screen "P_Bar_1" 1024x768
   Bar "Default" at 10,10 size 40x120
   TextField "Label_Default" at 10,132 size 51x20; Text 'Default'
   Bar "BackColor" at 60,10 size 40x120
   TextField "Label_BackColor" at 60,132 size 67x20; Text 'BackColor'
   Bar "BarBackColor" at 110,10 size 40x120
   TextField "Label_BarBackColor" at 110,132 size 89x20; Text 'BarBackColor'
   Bar "BarEdgeStyle" at 160,10 size 40x120
   TextField "Label_BarEdgeStyle" at 160,132 size 90x20; Text 'BarEdgeStyle'
   Bar "BarEdgeStyle_2" at 210,10 size 40x120
   TextField "Label_BarEdgeStyle_2" at 210,132 size 106x20; Text 'BarEdgeStyle_2'
   Bar "BarOrientation" at 260,10 size 40x120
   TextField "Label_BarOrientation" at 260,132 size 99x20; Text 'BarOrientation'
   Bar "BarOrientation_2" at 310,10 size 40x120
   TextField "Label_BarOrientation_2" at 310,132 size 115x20; Text 'BarOrientation_2'
   Bar "BarOrientation_3" at 360,10 size 40x120
   TextField "Label_BarOrientation_3" at 360,132 size 115x20; Text 'BarOrientation_3'
   Bar "BorderBackColor" at 410,10 size 40x120
   TextField "Label_BorderBackColor" at 410,132 size 111x20; Text 'BorderBackColor'
   Bar "BorderColor" at 460,10 size 40x120
   TextField "Label_BorderColor" at 460,132 size 81x20; Text 'BorderColor'
   Bar "BorderWidth" at 510,10 size 40x120
   TextField "Label_BorderWidth" at 510,132 size 86x20; Text 'BorderWidth'
   Bar "CornerRadius" at 560,10 size 40x120
   TextField "Label_CornerRadius" at 560,132 size 91x20; Text 'CornerRadius'
   Bar "CountSubDivisions" at 610,10 size 40x120
   TextField "Label_CountSubDivisions" at 610,132 size 122x20; Text 'CountSubDivisions'
   Bar "EdgeStyle" at 660,10 size 40x120
   TextField "Label_EdgeStyle" at 660,132 size 68x20; Text 'EdgeStyle'
   Bar "EdgeStyle_2" at 710,10 size 40x120
   TextField "Label_EdgeStyle_2" at 710,132 size 84x20; Text 'EdgeStyle_2'
   Bar "EdgeStyle_3" at 760,10 size 40x120
   TextField "Label_EdgeStyle_3" at 760,132 size 84x20; Text 'EdgeStyle_3'
   Bar "EdgeStyle_4" at 810,10 size 40x120
   TextField "Label_EdgeStyle_4" at 810,132 size 84x20; Text 'EdgeStyle_4'
   Bar "Flashing" at 860,10 size 40x120
   TextField "Label_Flashing" at 860,132 size 55x20; Text 'Flashing'
   Bar "FlashingOnLimitViolation" at 910,10 size 40x120
   TextField "Label_FlashingOnLimitViolation" at 910,132 size 158x20; Text 'FlashingOnLimitViolation'
   Bar "ForeColor" at 960,10 size 40x120
   TextField "Label_ForeColor" at 960,132 size 65x20; Text 'ForeColor'
   Bar "IntegerDigits" at 10,156 size 40x120
   TextField "Label_IntegerDigits" at 10,278 size 89x20; Text 'IntegerDigits'
   Bar "LargeTickLabelingStep" at 60,156 size 40x120
   TextField "Label_LargeTickLabelingStep" at 60,278 size 148x20; Text 'LargeTickLabelingStep'
   Bar "MaximumValue" at 110,156 size 40x120; MaximumValue 200
   TextField "Label_MaximumValue" at 110,278 size 99x20; Text 'MaximumValue'
   Bar "MinimumValue" at 160,156 size 40x120; MinimumValue -100
   TextField "Label_MinimumValue" at 160,278 size 95x20; Text 'MinimumValue'
   Bar "Precision" at 210,156 size 40x120
   TextField "Label_Precision" at 210,278 size 62x20; Text 'Precision'
   Bar "RangeLower1Color" at 260,156 size 40x120
   TextField "Label_RangeLower1Color" at 260,278 size 126x20; Text 'RangeLower1Color'
   Bar "RangeLower1Enabled" at 310,156 size 40x120
   TextField "Label_RangeLower1Enabled" at 310,278 size 143x20; Text 'RangeLower1Enabled'
   Bar "RangeLower2Color" at 360,156 size 40x120
   TextField "Label_RangeLower2Color" at 360,278 size 126x20; Text 'RangeLower2Color'
   Bar "RangeLower2Enabled" at 410,156 size 40x120
   TextField "Label_RangeLower2Enabled" at 410,278 size 143x20; Text 'RangeLower2Enabled'
   Bar "RangeNormalColor" at 460,156 size 40x120
   TextField "Label_RangeNormalColor" at 460,278 size 122x20; Text 'RangeNormalColor'
   Bar "RangeNormalEnabled" at 510,156 size 40x120
   TextField "Label_RangeNormalEnabled" at 510,278 size 139x20; Text 'RangeNormalEnabled'
   Bar "RangeUpper1Color" at 560,156 size 40x120
   TextField "Label_RangeUpper1Color" at 560,278 size 124x20; Text 'RangeUpper1Color'
   Bar "RangeUpper1Enabled" at 610,156 size 40x120
   TextField "Label_RangeUpper1Enabled" at 610,278 size 141x20; Text 'RangeUpper1Enabled'
   Bar "RangeUpper2Color" at 660,156 size 40x120
   TextField "Label_RangeUpper2Color" at 660,278 size 124x20; Text 'RangeUpper2Color'
   Bar "RangeUpper2Enabled" at 710,156 size 40x120
   TextField "Label_RangeUpper2Enabled" at 710,278 size 141x20; Text 'RangeUpper2Enabled'
   Bar "ScaleColor" at 760,156 size 40x120
   TextField "Label_ScaleColor" at 760,278 size 71x20; Text 'ScaleColor'
   Bar "ScaleGradation" at 810,156 size 40x120
   TextField "Label_ScaleGradation" at 810,278 size 101x20; Text 'ScaleGradation'
   Bar "ScaleLabelingDoubleLined" at 860,156 size 40x120
   TextField "Label_ScaleLabelingDoubleLined" at 860,278 size 169x20; Text 'ScaleLabelingDoubleLined'
   Bar "ScalePosition" at 910,156 size 40x120
   TextField "Label_ScalePosition" at 910,278 size 89x20; Text 'ScalePosition'
   Bar "SegmentColoring" at 960,156 size 40x120
   TextField "Label_SegmentColoring" at 960,278 size 113x20; Text 'SegmentColoring'
   Bar "ShowLimitLines" at 10,302 size 40x120
   TextField "Label_ShowLimitLines" at 10,424 size 102x20; Text 'ShowLimitLines'
   Bar "ShowLimitMarkers" at 60,302 size 40x120
   TextField "Label_ShowLimitMarkers" at 60,424 size 122x20; Text 'ShowLimitMarkers'
   Bar "ShowLimitRanges" at 110,302 size 40x120
   TextField "Label_ShowLimitRanges" at 110,424 size 117x20; Text 'ShowLimitRanges'
   Bar "ShowProcessValue" at 160,302 size 40x120
   TextField "Label_ShowProcessValue" at 160,424 size 126x20; Text 'ShowProcessValue'
   Bar "ShowScale" at 210,302 size 40x120
   TextField "Label_ShowScale" at 210,424 size 73x20; Text 'ShowScale'
   Bar "ShowTickLabels" at 260,302 size 40x120
   TextField "Label_ShowTickLabels" at 260,424 size 104x20; Text 'ShowTickLabels'
   Bar "Unit" at 310,302 size 40x120; Unit mm
   TextField "Label_Unit" at 310,424 size 29x20; Text 'Unit'
   Bar "UseAutoScaling" at 360,302 size 40x120
   TextField "Label_UseAutoScaling" at 360,424 size 104x20; Text 'UseAutoScaling'
   Bar "UseDesignColorSchema" at 410,302 size 40x120
   TextField "Label_UseDesignColorSchema" at 410,424 size 153x20; Text 'UseDesignColorSchema'
   Bar "UseExponentialFormat" at 460,302 size 40x120
   TextField "Label_UseExponentialFormat" at 460,424 size 146x20; Text 'UseExponentialFormat'
   Button "Next" at 982,744 size 40x22; TextOff 'Text'
      on Click: ActivateScreen("P_Switch_1", 0)

screen "P_Switch_1" 1024x768
   Switch "Default" at 10,10 size 120x40; CaptionText 'Switch'; TextOff '0'; TextOn '1'
   TextField "Label_Default" at 10,52 size 51x20; Text 'Default'
   Switch "AboveUpperLimitColor" at 140,10 size 120x40; CaptionText 'Switch'; TextOff '0'; TextOn '1'
   TextField "Label_AboveUpperLimitColor" at 140,52 size 147x20; Text 'AboveUpperLimitColor'
   Switch "BackColor" at 270,10 size 120x40; CaptionText 'Switch'; TextOff '0'; TextOn '1'
   TextField "Label_BackColor" at 270,52 size 67x20; Text 'BackColor'
   Switch "BackFillStyle" at 400,10 size 120x40; CaptionText 'Switch'; TextOff '0'; TextOn '1'
   TextField "Label_BackFillStyle" at 400,52 size 82x20; Text 'BackFillStyle'
   Switch "BelowLowerLimitColor" at 530,10 size 120x40; CaptionText 'Switch'; TextOff '0'; TextOn '1'
   TextField "Label_BelowLowerLimitColor" at 530,52 size 145x20; Text 'BelowLowerLimitColor'
   Switch "BorderBackColor" at 660,10 size 120x40; CaptionText 'Switch'; TextOff '0'; TextOn '1'
   TextField "Label_BorderBackColor" at 660,52 size 111x20; Text 'BorderBackColor'
   Switch "BorderColor" at 790,10 size 120x40; CaptionText 'Switch'; TextOff '0'; TextOn '1'
   TextField "Label_BorderColor" at 790,52 size 81x20; Text 'BorderColor'
   Switch "BorderWidth" at 10,76 size 120x40; CaptionText 'Switch'; TextOff '0'; TextOn '1'
   TextField "Label_BorderWidth" at 10,118 size 86x20; Text 'BorderWidth'
   Switch "CaptionColor" at 140,76 size 120x40; CaptionText 'Switch'; TextOff '0'; TextOn '1'
   TextField "Label_CaptionColor" at 140,118 size 86x20; Text 'CaptionColor'
   Switch "CornerRadius" at 270,76 size 120x40; CaptionText 'Switch'; TextOff '0'; TextOn '1'
   TextField "Label_CornerRadius" at 270,118 size 91x20; Text 'CornerRadius'
   Switch "EdgeStyle" at 400,76 size 120x40; CaptionText 'Switch'; TextOff '0'; TextOn '1'
   TextField "Label_EdgeStyle" at 400,118 size 68x20; Text 'EdgeStyle'
   Switch "EdgeStyle_2" at 530,76 size 120x40; CaptionText 'Switch'; TextOff '0'; TextOn '1'
   TextField "Label_EdgeStyle_2" at 530,118 size 84x20; Text 'EdgeStyle_2'
   Switch "EdgeStyle_3" at 660,76 size 120x40; CaptionText 'Switch'; TextOff '0'; TextOn '1'
   TextField "Label_EdgeStyle_3" at 660,118 size 84x20; Text 'EdgeStyle_3'
   Switch "EdgeStyle_4" at 790,76 size 120x40; CaptionText 'Switch'; TextOff '0'; TextOn '1'
   TextField "Label_EdgeStyle_4" at 790,118 size 84x20; Text 'EdgeStyle_4'
   Switch "FirstGradientColor" at 10,142 size 120x40; CaptionText 'Switch'; TextOff '0'; TextOn '1'
   TextField "Label_FirstGradientColor" at 10,184 size 120x20; Text 'FirstGradientColor'
   Switch "FirstGradientOffset" at 140,142 size 120x40; CaptionText 'Switch'; TextOff '0'; TextOn '1'
   TextField "Label_FirstGradientOffset" at 140,184 size 127x20; Text 'FirstGradientOffset'
   Switch "FitToLargest" at 270,142 size 120x40; CaptionText 'Switch'; TextOff '0'; TextOn '1'
   TextField "Label_FitToLargest" at 270,184 size 84x20; Text 'FitToLargest'
   Switch "Flashing" at 400,142 size 120x40; CaptionText 'Switch'; TextOff '0'; TextOn '1'
   TextField "Label_Flashing" at 400,184 size 55x20; Text 'Flashing'
   Switch "FlashingOnLimitViolation" at 530,142 size 120x40; CaptionText 'Switch'; TextOff '0'; TextOn '1'
   TextField "Label_FlashingOnLimitViolation" at 530,184 size 158x20; Text 'FlashingOnLimitViolation'
   Switch "FocusColor" at 660,142 size 120x40; CaptionText 'Switch'; TextOff '0'; TextOn '1'
   TextField "Label_FocusColor" at 660,184 size 73x20; Text 'FocusColor'
   Switch "FocusWidth" at 790,142 size 120x40; CaptionText 'Switch'; TextOff '0'; TextOn '1'
   TextField "Label_FocusWidth" at 790,184 size 78x20; Text 'FocusWidth'
   Switch "ForeColor" at 10,208 size 120x40; CaptionText 'Switch'; TextOff '0'; TextOn '1'
   TextField "Label_ForeColor" at 10,250 size 65x20; Text 'ForeColor'
   Switch "HorizontalAlignment" at 140,208 size 120x40; CaptionText 'Switch'; TextOff '0'; TextOn '1'
   TextField "Label_HorizontalAlignment" at 140,250 size 135x20; Text 'HorizontalAlignment'
   Switch "HorizontalAlignment_2" at 270,208 size 120x40; CaptionText 'Switch'; TextOff '0'; TextOn '1'
   TextField "Label_HorizontalAlignment_2" at 270,250 size 151x20; Text 'HorizontalAlignment_2'
   Switch "HorizontalPictureAlignment" at 400,208 size 120x40; CaptionText 'Switch'; TextOff '0'; TextOn '1'
   TextField "Label_HorizontalPictureAlignment" at 400,250 size 181x20; Text 'HorizontalPictureAlignment'
   Switch "HorizontalPictureAlignment_2" at 530,208 size 120x40; CaptionText 'Switch'; TextOff '0'; TextOn '1'
   TextField "Label_HorizontalPictureAlignment_2" at 530,250 size 197x20; Text 'HorizontalPictureAlignment_2'
   Switch "InnerBackColorOff" at 660,208 size 120x40; CaptionText 'Switch'; TextOff '0'; TextOn '1'
   TextField "Label_InnerBackColorOff" at 660,250 size 121x20; Text 'InnerBackColorOff'
   Switch "InnerBackColorOn" at 790,208 size 120x40; CaptionText 'Switch'; TextOff '0'; TextOn '1'
   TextField "Label_InnerBackColorOn" at 790,250 size 119x20; Text 'InnerBackColorOn'
   Switch "MiddleGradientColor" at 10,274 size 120x40; CaptionText 'Switch'; TextOff '0'; TextOn '1'
   TextField "Label_MiddleGradientColor" at 10,316 size 133x20; Text 'MiddleGradientColor'
   Switch "PictureAreaBottomMargin" at 140,274 size 120x40; CaptionText 'Switch'; TextOff '0'; TextOn '1'
   TextField "Label_PictureAreaBottomMargin" at 140,316 size 173x20; Text 'PictureAreaBottomMargin'
   Switch "PictureAreaLeftMargin" at 270,274 size 120x40; CaptionText 'Switch'; TextOff '0'; TextOn '1'
   TextField "Label_PictureAreaLeftMargin" at 270,316 size 152x20; Text 'PictureAreaLeftMargin'
   Switch "PictureAreaRightMargin" at 400,274 size 120x40; CaptionText 'Switch'; TextOff '0'; TextOn '1'
   TextField "Label_PictureAreaRightMargin" at 400,316 size 160x20; Text 'PictureAreaRightMargin'
   Switch "PictureAreaTopMargin" at 530,274 size 120x40; CaptionText 'Switch'; TextOff '0'; TextOn '1'
   TextField "Label_PictureAreaTopMargin" at 530,316 size 149x20; Text 'PictureAreaTopMargin'
   Switch "SecondGradientColor" at 660,274 size 120x40; CaptionText 'Switch'; TextOff '0'; TextOn '1'
   TextField "Label_SecondGradientColor" at 660,316 size 139x20; Text 'SecondGradientColor'
   Switch "SecondGradientOffset" at 790,274 size 120x40; CaptionText 'Switch'; TextOff '0'; TextOn '1'
   TextField "Label_SecondGradientOffset" at 790,316 size 146x20; Text 'SecondGradientOffset'
   Switch "ShowCaption" at 10,340 size 120x40; CaptionText 'Switch'; TextOff '0'; TextOn '1'
   TextField "Label_ShowCaption" at 10,382 size 88x20; Text 'ShowCaption'
   Switch "SwitchOrientation" at 140,340 size 120x40; CaptionText 'Switch'; TextOff '0'; TextOn '1'
   TextField "Label_SwitchOrientation" at 140,382 size 120x20; Text 'SwitchOrientation'
   Switch "SwitchOrientation_2" at 270,340 size 120x40; CaptionText 'Switch'; TextOff '0'; TextOn '1'
   TextField "Label_SwitchOrientation_2" at 270,382 size 136x20; Text 'SwitchOrientation_2'
   Switch "SwitchOrientation_3" at 400,340 size 120x40; CaptionText 'Switch'; TextOff '0'; TextOn '1'
   TextField "Label_SwitchOrientation_3" at 400,382 size 136x20; Text 'SwitchOrientation_3'
   Switch "TextAreaBottomMargin" at 530,340 size 120x40; CaptionText 'Switch'; TextOff '0'; TextOn '1'
   TextField "Label_TextAreaBottomMargin" at 530,382 size 155x20; Text 'TextAreaBottomMargin'
   Switch "TextAreaLeftMargin" at 660,340 size 120x40; CaptionText 'Switch'; TextOff '0'; TextOn '1'
   TextField "Label_TextAreaLeftMargin" at 660,382 size 134x20; Text 'TextAreaLeftMargin'
   Switch "TextAreaRightMargin" at 790,340 size 120x40; CaptionText 'Switch'; TextOff '0'; TextOn '1'
   TextField "Label_TextAreaRightMargin" at 790,382 size 142x20; Text 'TextAreaRightMargin'
   Switch "TextAreaTopMargin" at 10,406 size 120x40; CaptionText 'Switch'; TextOff '0'; TextOn '1'
   TextField "Label_TextAreaTopMargin" at 10,448 size 131x20; Text 'TextAreaTopMargin'
   Switch "UseDesignColorSchema" at 140,406 size 120x40; CaptionText 'Switch'; TextOff '0'; TextOn '1'
   TextField "Label_UseDesignColorSchema" at 140,448 size 153x20; Text 'UseDesignColorSchema'
   Switch "UseFirstGradient" at 270,406 size 120x40; CaptionText 'Switch'; TextOff '0'; TextOn '1'
   TextField "Label_UseFirstGradient" at 270,448 size 110x20; Text 'UseFirstGradient'
   Switch "UseSecondGradient" at 400,406 size 120x40; CaptionText 'Switch'; TextOff '0'; TextOn '1'
   TextField "Label_UseSecondGradient" at 400,448 size 129x20; Text 'UseSecondGradient'
   Switch "VerticalAlignment" at 530,406 size 120x40; CaptionText 'Switch'; TextOff '0'; TextOn '1'
   TextField "Label_VerticalAlignment" at 530,448 size 119x20; Text 'VerticalAlignment'
   Switch "VerticalAlignment_2" at 660,406 size 120x40; CaptionText 'Switch'; TextOff '0'; TextOn '1'
   TextField "Label_VerticalAlignment_2" at 660,448 size 135x20; Text 'VerticalAlignment_2'
   Switch "VerticalPictureAlignment" at 790,406 size 120x40; CaptionText 'Switch'; TextOff '0'; TextOn '1'
   TextField "Label_VerticalPictureAlignment" at 790,448 size 165x20; Text 'VerticalPictureAlignment'
   Switch "VerticalPictureAlignment_2" at 10,472 size 120x40; CaptionText 'Switch'; TextOff '0'; TextOn '1'
   TextField "Label_VerticalPictureAlignment_2" at 10,514 size 181x20; Text 'VerticalPictureAlignment_2'
   Button "Next" at 982,744 size 40x22; TextOff 'Text'
      on Click: ActivateScreen("P_SymbolLibrary_1", 0)

screen "P_SymbolLibrary_1" 1024x768
   SymbolLibrary "Default" at 10,10 size 60x60
   TextField "Label_Default" at 10,72 size 51x20; Text 'Default'
   SymbolLibrary "AboveUpperLimitColor" at 80,10 size 60x60
   TextField "Label_AboveUpperLimitColor" at 80,72 size 147x20; Text 'AboveUpperLimitColor'
   SymbolLibrary "BackColor" at 150,10 size 60x60
   TextField "Label_BackColor" at 150,72 size 67x20; Text 'BackColor'
   SymbolLibrary "BackFillStyle" at 220,10 size 60x60
   TextField "Label_BackFillStyle" at 220,72 size 82x20; Text 'BackFillStyle'
   SymbolLibrary "BelowLowerLimitColor" at 290,10 size 60x60
   TextField "Label_BelowLowerLimitColor" at 290,72 size 145x20; Text 'BelowLowerLimitColor'
   SymbolLibrary "BlinkColor" at 360,10 size 60x60
   TextField "Label_BlinkColor" at 360,72 size 66x20; Text 'BlinkColor'
   SymbolLibrary "FillColorMode" at 430,10 size 60x60
   TextField "Label_FillColorMode" at 430,72 size 87x20; Text 'FillColorMode'
   SymbolLibrary "FillColorMode_2" at 500,10 size 60x60
   TextField "Label_FillColorMode_2" at 500,72 size 103x20; Text 'FillColorMode_2'
   SymbolLibrary "FixedAspectRatio" at 570,10 size 60x60
   TextField "Label_FixedAspectRatio" at 570,72 size 116x20; Text 'FixedAspectRatio'
   SymbolLibrary "Flashing" at 640,10 size 60x60
   TextField "Label_Flashing" at 640,72 size 55x20; Text 'Flashing'
   SymbolLibrary "FlashingOnLimitViolation" at 710,10 size 60x60
   TextField "Label_FlashingOnLimitViolation" at 710,72 size 158x20; Text 'FlashingOnLimitViolation'
   SymbolLibrary "Flip" at 780,10 size 60x60
   TextField "Label_Flip" at 780,72 size 24x20; Text 'Flip'
   SymbolLibrary "Flip_2" at 850,10 size 60x60
   TextField "Label_Flip_2" at 850,72 size 40x20; Text 'Flip_2'
   SymbolLibrary "Flip_3" at 920,10 size 60x60
   TextField "Label_Flip_3" at 920,72 size 40x20; Text 'Flip_3'
   SymbolLibrary "ForeColor" at 10,96 size 60x60
   TextField "Label_ForeColor" at 10,158 size 65x20; Text 'ForeColor'
   SymbolLibrary "Rotation" at 80,96 size 60x60
   TextField "Label_Rotation" at 80,158 size 60x20; Text 'Rotation'
   SymbolLibrary "Rotation_2" at 150,96 size 60x60
   TextField "Label_Rotation_2" at 150,158 size 76x20; Text 'Rotation_2'
   SymbolLibrary "Rotation_3" at 220,96 size 60x60
   TextField "Label_Rotation_3" at 220,158 size 76x20; Text 'Rotation_3'
   Button "Next" at 982,744 size 40x22; TextOff 'Text'
      on Click: ActivateScreen("P_Slider_1", 0)

screen "P_Slider_1" 1024x768
   Slider "Default" at 10,10 size 60x160; Caption 'SIMATIC'
   TextField "Label_Default" at 10,172 size 51x20; Text 'Default'
   Slider "BackColor" at 80,10 size 60x160; Caption 'SIMATIC'
   TextField "Label_BackColor" at 80,172 size 67x20; Text 'BackColor'
   Slider "BackFillStyle" at 150,10 size 60x160; Caption 'SIMATIC'
   TextField "Label_BackFillStyle" at 150,172 size 82x20; Text 'BackFillStyle'
   Slider "BarBackColor" at 220,10 size 60x160; Caption 'SIMATIC'
   TextField "Label_BarBackColor" at 220,172 size 89x20; Text 'BarBackColor'
   Slider "BarColor" at 290,10 size 60x160; Caption 'SIMATIC'
   TextField "Label_BarColor" at 290,172 size 59x20; Text 'BarColor'
   Slider "BarOrientation" at 360,10 size 60x160; Caption 'SIMATIC'
   TextField "Label_BarOrientation" at 360,172 size 99x20; Text 'BarOrientation'
   Slider "BarOrientation_2" at 430,10 size 60x160; Caption 'SIMATIC'
   TextField "Label_BarOrientation_2" at 430,172 size 115x20; Text 'BarOrientation_2'
   Slider "BarOrientation_3" at 500,10 size 60x160; Caption 'SIMATIC'
   TextField "Label_BarOrientation_3" at 500,172 size 115x20; Text 'BarOrientation_3'
   Slider "BorderBackColor" at 570,10 size 60x160; Caption 'SIMATIC'
   TextField "Label_BorderBackColor" at 570,172 size 111x20; Text 'BorderBackColor'
   Slider "BorderBrightColor3D" at 640,10 size 60x160; Caption 'SIMATIC'
   TextField "Label_BorderBrightColor3D" at 640,172 size 137x20; Text 'BorderBrightColor3D'
   Slider "BorderColor" at 710,10 size 60x160; Caption 'SIMATIC'
   TextField "Label_BorderColor" at 710,172 size 81x20; Text 'BorderColor'
   Slider "BorderInnerStyle3D" at 780,10 size 60x160; Caption 'SIMATIC'
   TextField "Label_BorderInnerStyle3D" at 780,172 size 133x20; Text 'BorderInnerStyle3D'
   Slider "BorderInnerStyle3D_2" at 850,10 size 60x160; Caption 'SIMATIC'
   TextField "Label_BorderInnerStyle3D_2" at 850,172 size 149x20; Text 'BorderInnerStyle3D_2'
   Slider "BorderInnerWidth3D" at 920,10 size 60x160; Caption 'SIMATIC'
   TextField "Label_BorderInnerWidth3D" at 920,172 size 138x20; Text 'BorderInnerWidth3D'
   Slider "BorderOuterStyle3D" at 10,196 size 60x160; Caption 'SIMATIC'
   TextField "Label_BorderOuterStyle3D" at 10,358 size 135x20; Text 'BorderOuterStyle3D'
   Slider "BorderOuterStyle3D_2" at 80,196 size 60x160; Caption 'SIMATIC'
   TextField "Label_BorderOuterStyle3D_2" at 80,358 size 151x20; Text 'BorderOuterStyle3D_2'
   Slider "BorderOuterWidth3D" at 150,196 size 60x160; Caption 'SIMATIC'
   TextField "Label_BorderOuterWidth3D" at 150,358 size 140x20; Text 'BorderOuterWidth3D'
   Slider "BorderShadeColor3D" at 220,196 size 60x160; Caption 'SIMATIC'
   TextField "Label_BorderShadeColor3D" at 220,358 size 138x20; Text 'BorderShadeColor3D'
   Slider "BorderWidth" at 290,196 size 60x160; Caption 'SIMATIC'
   TextField "Label_BorderWidth" at 290,358 size 86x20; Text 'BorderWidth'
   Slider "CornerRadius" at 360,196 size 60x160; Caption 'SIMATIC'
   TextField "Label_CornerRadius" at 360,358 size 91x20; Text 'CornerRadius'
   Slider "EdgeStyle" at 430,196 size 60x160; Caption 'SIMATIC'
   TextField "Label_EdgeStyle" at 430,358 size 68x20; Text 'EdgeStyle'
   Slider "EdgeStyle_2" at 500,196 size 60x160; Caption 'SIMATIC'
   TextField "Label_EdgeStyle_2" at 500,358 size 84x20; Text 'EdgeStyle_2'
   Slider "EdgeStyle_3" at 570,196 size 60x160; Caption 'SIMATIC'
   TextField "Label_EdgeStyle_3" at 570,358 size 84x20; Text 'EdgeStyle_3'
   Slider "EdgeStyle_4" at 640,196 size 60x160; Caption 'SIMATIC'
   TextField "Label_EdgeStyle_4" at 640,358 size 84x20; Text 'EdgeStyle_4'
   Slider "Flashing" at 710,196 size 60x160; Caption 'SIMATIC'
   TextField "Label_Flashing" at 710,358 size 55x20; Text 'Flashing'
   Slider "FocusColor" at 780,196 size 60x160; Caption 'SIMATIC'
   TextField "Label_FocusColor" at 780,358 size 73x20; Text 'FocusColor'
   Slider "FocusWidth" at 850,196 size 60x160; Caption 'SIMATIC'
   TextField "Label_FocusWidth" at 850,358 size 78x20; Text 'FocusWidth'
   Slider "ForeColor" at 920,196 size 60x160; Caption 'SIMATIC'
   TextField "Label_ForeColor" at 920,358 size 65x20; Text 'ForeColor'
   Slider "LabelColor" at 10,382 size 60x160; Caption 'SIMATIC'
   TextField "Label_LabelColor" at 10,544 size 71x20; Text 'LabelColor'
   Slider "MaximumValue" at 80,382 size 60x160; Caption 'SIMATIC'
   TextField "Label_MaximumValue" at 80,544 size 99x20; Text 'MaximumValue'
   Slider "MinimumValue" at 150,382 size 60x160; Caption 'SIMATIC'
   TextField "Label_MinimumValue" at 150,544 size 95x20; Text 'MinimumValue'
   Slider "RangeLower1Color" at 220,382 size 60x160; Caption 'SIMATIC'
   TextField "Label_RangeLower1Color" at 220,544 size 126x20; Text 'RangeLower1Color'
   Slider "RangeLower1Enabled" at 290,382 size 60x160; Caption 'SIMATIC'
   TextField "Label_RangeLower1Enabled" at 290,544 size 143x20; Text 'RangeLower1Enabled'
   Slider "RangeLower2Color" at 360,382 size 60x160; Caption 'SIMATIC'
   TextField "Label_RangeLower2Color" at 360,544 size 126x20; Text 'RangeLower2Color'
   Slider "RangeLower2Enabled" at 430,382 size 60x160; Caption 'SIMATIC'
   TextField "Label_RangeLower2Enabled" at 430,544 size 143x20; Text 'RangeLower2Enabled'
   Slider "RangeNormalColor" at 500,382 size 60x160; Caption 'SIMATIC'
   TextField "Label_RangeNormalColor" at 500,544 size 122x20; Text 'RangeNormalColor'
   Slider "RangeNormalEnabled" at 570,382 size 60x160; Caption 'SIMATIC'
   TextField "Label_RangeNormalEnabled" at 570,544 size 139x20; Text 'RangeNormalEnabled'
   Slider "RangeUpper1Color" at 640,382 size 60x160; Caption 'SIMATIC'
   TextField "Label_RangeUpper1Color" at 640,544 size 124x20; Text 'RangeUpper1Color'
   Slider "RangeUpper1Enabled" at 710,382 size 60x160; Caption 'SIMATIC'
   TextField "Label_RangeUpper1Enabled" at 710,544 size 141x20; Text 'RangeUpper1Enabled'
   Slider "RangeUpper2Color" at 780,382 size 60x160; Caption 'SIMATIC'
   TextField "Label_RangeUpper2Color" at 780,544 size 124x20; Text 'RangeUpper2Color'
   Slider "RangeUpper2Enabled" at 850,382 size 60x160; Caption 'SIMATIC'
   TextField "Label_RangeUpper2Enabled" at 850,544 size 141x20; Text 'RangeUpper2Enabled'
   Slider "ScalePosition" at 920,382 size 60x160; Caption 'SIMATIC'
   TextField "Label_ScalePosition" at 920,544 size 89x20; Text 'ScalePosition'
   Button "Next" at 982,744 size 40x22; TextOff 'Text'
      on Click: ActivateScreen("P_Slider_2", 0)

screen "P_Slider_2" 1024x768
   Slider "ShowBar" at 10,10 size 60x160; Caption 'SIMATIC'
   TextField "Label_ShowBar" at 10,172 size 61x20; Text 'ShowBar'
   Slider "ShowLimitLines" at 80,10 size 60x160; Caption 'SIMATIC'
   TextField "Label_ShowLimitLines" at 80,172 size 102x20; Text 'ShowLimitLines'
   Slider "ShowLimitMarkers" at 150,10 size 60x160; Caption 'SIMATIC'
   TextField "Label_ShowLimitMarkers" at 150,172 size 122x20; Text 'ShowLimitMarkers'
   Slider "ShowLimitRanges" at 220,10 size 60x160; Caption 'SIMATIC'
   TextField "Label_ShowLimitRanges" at 220,172 size 117x20; Text 'ShowLimitRanges'
   Slider "ShowPosition" at 290,10 size 60x160; Caption 'SIMATIC'
   TextField "Label_ShowPosition" at 290,172 size 90x20; Text 'ShowPosition'
   Slider "ShowScale" at 360,10 size 60x160; Caption 'SIMATIC'
   TextField "Label_ShowScale" at 360,172 size 73x20; Text 'ShowScale'
   Slider "ShowThumb" at 430,10 size 60x160; Caption 'SIMATIC'
   TextField "Label_ShowThumb" at 430,172 size 81x20; Text 'ShowThumb'
   Slider "ShowTickLabels" at 500,10 size 60x160; Caption 'SIMATIC'
   TextField "Label_ShowTickLabels" at 500,172 size 104x20; Text 'ShowTickLabels'
   Slider "ShowTicks" at 570,10 size 60x160; Caption 'SIMATIC'
   TextField "Label_ShowTicks" at 570,172 size 70x20; Text 'ShowTicks'
   Slider "ThumbBackColor" at 640,10 size 60x160; Caption 'SIMATIC'
   TextField "Label_ThumbBackColor" at 640,172 size 109x20; Text 'ThumbBackColor'
   Slider "UseDesignColorSchema" at 710,10 size 60x160; Caption 'SIMATIC'
   TextField "Label_UseDesignColorSchema" at 710,172 size 153x20; Text 'UseDesignColorSchema'
   Button "Next" at 982,744 size 40x22; TextOff 'Text'
      on Click: ActivateScreen("P_Gauge_1", 0)

screen "P_Gauge_1" 1024x768
   Gauge "Default" at 10,10 size 150x150; CaptionText 'SIMATIC'
   TextField "Label_Default" at 10,162 size 51x20; Text 'Default'
   Gauge "AngleMax" at 170,10 size 150x150; CaptionText 'SIMATIC'
   TextField "Label_AngleMax" at 170,162 size 67x20; Text 'AngleMax'
   Gauge "AngleMin" at 330,10 size 150x150; CaptionText 'SIMATIC'
   TextField "Label_AngleMin" at 330,162 size 63x20; Text 'AngleMin'
   Gauge "BackColor" at 490,10 size 150x150; CaptionText 'SIMATIC'
   TextField "Label_BackColor" at 490,162 size 67x20; Text 'BackColor'
   Gauge "BackFillStyle" at 650,10 size 150x150; CaptionText 'SIMATIC'
   TextField "Label_BackFillStyle" at 650,162 size 82x20; Text 'BackFillStyle'
   Gauge "BorderBackColor" at 810,10 size 150x150; CaptionText 'SIMATIC'
   TextField "Label_BorderBackColor" at 810,162 size 111x20; Text 'BorderBackColor'
   Gauge "BorderColor" at 10,186 size 150x150; CaptionText 'SIMATIC'
   TextField "Label_BorderColor" at 10,338 size 81x20; Text 'BorderColor'
   Gauge "BorderWidth" at 170,186 size 150x150; CaptionText 'SIMATIC'
   TextField "Label_BorderWidth" at 170,338 size 86x20; Text 'BorderWidth'
   Gauge "CaptionColor" at 330,186 size 150x150; CaptionText 'SIMATIC'
   TextField "Label_CaptionColor" at 330,338 size 86x20; Text 'CaptionColor'
   Gauge "CaptionTop" at 490,186 size 150x150; CaptionText 'SIMATIC'
   TextField "Label_CaptionTop" at 490,338 size 76x20; Text 'CaptionTop'
   Gauge "CenterColor" at 650,186 size 150x150; CaptionText 'SIMATIC'
   TextField "Label_CenterColor" at 650,338 size 81x20; Text 'CenterColor'
   Gauge "CenterSize" at 810,186 size 150x150; CaptionText 'SIMATIC'
   TextField "Label_CenterSize" at 810,338 size 74x20; Text 'CenterSize'
   Gauge "CornerRadius" at 10,362 size 150x150; CaptionText 'SIMATIC'
   TextField "Label_CornerRadius" at 10,514 size 91x20; Text 'CornerRadius'
   Gauge "DialColor" at 170,362 size 150x150; CaptionText 'SIMATIC'
   TextField "Label_DialColor" at 170,514 size 60x20; Text 'DialColor'
   Gauge "DialFillStyle" at 330,362 size 150x150; CaptionText 'SIMATIC'
   TextField "Label_DialFillStyle" at 330,514 size 75x20; Text 'DialFillStyle'
   Gauge "DialSize" at 490,362 size 150x150; CaptionText 'SIMATIC'
   TextField "Label_DialSize" at 490,514 size 53x20; Text 'DialSize'
   Gauge "EdgeStyle" at 650,362 size 150x150; CaptionText 'SIMATIC'
   TextField "Label_EdgeStyle" at 650,514 size 68x20; Text 'EdgeStyle'
   Gauge "EdgeStyle_2" at 810,362 size 150x150; CaptionText 'SIMATIC'
   TextField "Label_EdgeStyle_2" at 810,514 size 84x20; Text 'EdgeStyle_2'
   Gauge "EdgeStyle_3" at 10,538 size 150x150; CaptionText 'SIMATIC'
   TextField "Label_EdgeStyle_3" at 10,690 size 84x20; Text 'EdgeStyle_3'
   Gauge "EdgeStyle_4" at 170,538 size 150x150; CaptionText 'SIMATIC'
   TextField "Label_EdgeStyle_4" at 170,690 size 84x20; Text 'EdgeStyle_4'
   Gauge "Gradation" at 330,538 size 150x150; CaptionText 'SIMATIC'
   TextField "Label_Gradation" at 330,690 size 67x20; Text 'Gradation'
   Gauge "InnerDialColor" at 490,538 size 150x150; CaptionText 'SIMATIC'
   TextField "Label_InnerDialColor" at 490,690 size 95x20; Text 'InnerDialColor'
   Gauge "InnerDialInnerDistance" at 650,538 size 150x150; CaptionText 'SIMATIC'
   TextField "Label_InnerDialInnerDistance" at 650,690 size 153x20; Text 'InnerDialInnerDistance'
   Gauge "InnerDialOuterDistance" at 810,538 size 150x150; CaptionText 'SIMATIC'
   TextField "Label_InnerDialOuterDistance" at 810,690 size 155x20; Text 'InnerDialOuterDistance'
   Button "Next" at 982,744 size 40x22; TextOff 'Text'
      on Click: ActivateScreen("P_Gauge_2", 0)

screen "P_Gauge_2" 1024x768
   Gauge "LockSquaredExtent" at 10,10 size 150x150; CaptionText 'SIMATIC'
   TextField "Label_LockSquaredExtent" at 10,162 size 129x20; Text 'LockSquaredExtent'
   Gauge "MaximumValue" at 170,10 size 150x150; CaptionText 'SIMATIC'
   TextField "Label_MaximumValue" at 170,162 size 99x20; Text 'MaximumValue'
   Gauge "MinimumValue" at 330,10 size 150x150; CaptionText 'SIMATIC'
   TextField "Label_MinimumValue" at 330,162 size 95x20; Text 'MinimumValue'
   Gauge "NeedleHeight" at 490,10 size 150x150; CaptionText 'SIMATIC'
   TextField "Label_NeedleHeight" at 490,162 size 89x20; Text 'NeedleHeight'
   Gauge "PointerColor" at 650,10 size 150x150; CaptionText 'SIMATIC'
   TextField "Label_PointerColor" at 650,162 size 84x20; Text 'PointerColor'
   Gauge "RangeLower1Color" at 810,10 size 150x150; CaptionText 'SIMATIC'
   TextField "Label_RangeLower1Color" at 810,162 size 126x20; Text 'RangeLower1Color'
   Gauge "RangeLower1Enabled" at 10,186 size 150x150; CaptionText 'SIMATIC'
   TextField "Label_RangeLower1Enabled" at 10,338 size 143x20; Text 'RangeLower1Enabled'
   Gauge "RangeLower2Color" at 170,186 size 150x150; CaptionText 'SIMATIC'
   TextField "Label_RangeLower2Color" at 170,338 size 126x20; Text 'RangeLower2Color'
   Gauge "RangeLower2Enabled" at 330,186 size 150x150; CaptionText 'SIMATIC'
   TextField "Label_RangeLower2Enabled" at 330,338 size 143x20; Text 'RangeLower2Enabled'
   Gauge "RangeNormalColor" at 490,186 size 150x150; CaptionText 'SIMATIC'
   TextField "Label_RangeNormalColor" at 490,338 size 122x20; Text 'RangeNormalColor'
   Gauge "RangeNormalEnabled" at 650,186 size 150x150; CaptionText 'SIMATIC'
   TextField "Label_RangeNormalEnabled" at 650,338 size 139x20; Text 'RangeNormalEnabled'
   Gauge "RangeUpper1Color" at 810,186 size 150x150; CaptionText 'SIMATIC'
   TextField "Label_RangeUpper1Color" at 810,338 size 124x20; Text 'RangeUpper1Color'
   Gauge "RangeUpper1Enabled" at 10,362 size 150x150; CaptionText 'SIMATIC'
   TextField "Label_RangeUpper1Enabled" at 10,514 size 141x20; Text 'RangeUpper1Enabled'
   Gauge "RangeUpper1Start" at 170,362 size 150x150; CaptionText 'SIMATIC'
   TextField "Label_RangeUpper1Start" at 170,514 size 125x20; Text 'RangeUpper1Start'
   Gauge "RangeUpper2Color" at 330,362 size 150x150; CaptionText 'SIMATIC'
   TextField "Label_RangeUpper2Color" at 330,514 size 124x20; Text 'RangeUpper2Color'
   Gauge "RangeUpper2Enabled" at 490,362 size 150x150; CaptionText 'SIMATIC'
   TextField "Label_RangeUpper2Enabled" at 490,514 size 141x20; Text 'RangeUpper2Enabled'
   Gauge "RangeUpper2Start" at 650,362 size 150x150; CaptionText 'SIMATIC'
   TextField "Label_RangeUpper2Start" at 650,514 size 125x20; Text 'RangeUpper2Start'
   Gauge "ScaleLabelColor" at 810,362 size 150x150; CaptionText 'SIMATIC'
   TextField "Label_ScaleLabelColor" at 810,514 size 105x20; Text 'ScaleLabelColor'
   Gauge "ScaleTickColor" at 10,538 size 150x150; CaptionText 'SIMATIC'
   TextField "Label_ScaleTickColor" at 10,690 size 95x20; Text 'ScaleTickColor'
   Gauge "ScaleTickLabelPosition" at 170,538 size 150x150; CaptionText 'SIMATIC'
   TextField "Label_ScaleTickLabelPosition" at 170,690 size 147x20; Text 'ScaleTickLabelPosition'
   Gauge "ScaleTickLength" at 330,538 size 150x150; CaptionText 'SIMATIC'
   TextField "Label_ScaleTickLength" at 330,690 size 107x20; Text 'ScaleTickLength'
   Gauge "ScaleTickPosition" at 490,538 size 150x150; CaptionText 'SIMATIC'
   TextField "Label_ScaleTickPosition" at 490,690 size 113x20; Text 'ScaleTickPosition'
   Gauge "ShowDecimalPoint" at 650,538 size 150x150; CaptionText 'SIMATIC'
   TextField "Label_ShowDecimalPoint" at 650,690 size 121x20; Text 'ShowDecimalPoint'
   Gauge "ShowInnerDial" at 810,538 size 150x150; CaptionText 'SIMATIC'
   TextField "Label_ShowInnerDial" at 810,690 size 97x20; Text 'ShowInnerDial'
   Button "Next" at 982,744 size 40x22; TextOff 'Text'
      on Click: ActivateScreen("P_Gauge_3", 0)

screen "P_Gauge_3" 1024x768
   Gauge "ShowLimitRanges" at 10,10 size 150x150; CaptionText 'SIMATIC'
   TextField "Label_ShowLimitRanges" at 10,162 size 117x20; Text 'ShowLimitRanges'
   Gauge "ShowPeakValuePointer" at 170,10 size 150x150; CaptionText 'SIMATIC'
   TextField "Label_ShowPeakValuePointer" at 170,162 size 153x20; Text 'ShowPeakValuePointer'
   Gauge "UnitColor" at 330,10 size 150x150; CaptionText 'SIMATIC'
   TextField "Label_UnitColor" at 330,162 size 62x20; Text 'UnitColor'
   Gauge "UnitTop" at 490,10 size 150x150; CaptionText 'SIMATIC'
   TextField "Label_UnitTop" at 490,162 size 52x20; Text 'UnitTop'
   Gauge "UseDesignColorSchema" at 650,10 size 150x150; CaptionText 'SIMATIC'
   TextField "Label_UseDesignColorSchema" at 650,162 size 153x20; Text 'UseDesignColorSchema'
   Button "Next" at 982,744 size 40x22; TextOff 'Text'
      on Click: ActivateScreen("P_Clock_1", 0)

screen "P_Clock_1" 1024x768
   Clock "Default" at 10,10 size 150x150
   TextField "Label_Default" at 10,162 size 51x20; Text 'Default'
   Clock "Analog" at 170,10 size 150x150
   TextField "Label_Analog" at 170,162 size 49x20; Text 'Analog'
   Clock "BackFillStyle" at 330,10 size 150x150
   TextField "Label_BackFillStyle" at 330,162 size 82x20; Text 'BackFillStyle'
   Clock "BorderBackColor" at 490,10 size 150x150
   TextField "Label_BorderBackColor" at 490,162 size 111x20; Text 'BorderBackColor'
   Clock "BorderColor" at 650,10 size 150x150
   TextField "Label_BorderColor" at 650,162 size 81x20; Text 'BorderColor'
   Clock "BorderWidth" at 810,10 size 150x150
   TextField "Label_BorderWidth" at 810,162 size 86x20; Text 'BorderWidth'
   Clock "CornerRadius" at 10,186 size 150x150
   TextField "Label_CornerRadius" at 10,338 size 91x20; Text 'CornerRadius'
   Clock "DialColor" at 170,186 size 150x150
   TextField "Label_DialColor" at 170,338 size 60x20; Text 'DialColor'
   Clock "EdgeStyle" at 330,186 size 150x150
   TextField "Label_EdgeStyle" at 330,338 size 68x20; Text 'EdgeStyle'
   Clock "EdgeStyle_2" at 490,186 size 150x150
   TextField "Label_EdgeStyle_2" at 490,338 size 84x20; Text 'EdgeStyle_2'
   Clock "EdgeStyle_3" at 650,186 size 150x150
   TextField "Label_EdgeStyle_3" at 650,338 size 84x20; Text 'EdgeStyle_3'
   Clock "EdgeStyle_4" at 810,186 size 150x150
   TextField "Label_EdgeStyle_4" at 810,338 size 84x20; Text 'EdgeStyle_4'
   Clock "Flashing" at 10,362 size 150x150
   TextField "Label_Flashing" at 10,514 size 55x20; Text 'Flashing'
   Clock "HourNeedleHeight" at 170,362 size 150x150
   TextField "Label_HourNeedleHeight" at 170,514 size 120x20; Text 'HourNeedleHeight'
   Clock "HourNeedleWidth" at 330,362 size 150x150
   TextField "Label_HourNeedleWidth" at 330,514 size 116x20; Text 'HourNeedleWidth'
   Clock "LockSquaredExtent" at 490,362 size 150x150
   TextField "Label_LockSquaredExtent" at 490,514 size 129x20; Text 'LockSquaredExtent'
   Clock "MinuteNeedleHeight" at 650,362 size 150x150
   TextField "Label_MinuteNeedleHeight" at 650,514 size 133x20; Text 'MinuteNeedleHeight'
   Clock "MinuteNeedleWidth" at 810,362 size 150x150
   TextField "Label_MinuteNeedleWidth" at 810,514 size 129x20; Text 'MinuteNeedleWidth'
   Clock "NeedleBorderColor" at 10,538 size 150x150
   TextField "Label_NeedleBorderColor" at 10,690 size 124x20; Text 'NeedleBorderColor'
   Clock "NeedleColor" at 170,538 size 150x150
   TextField "Label_NeedleColor" at 170,690 size 80x20; Text 'NeedleColor'
   Clock "NeedleFillStyle" at 330,538 size 150x150
   TextField "Label_NeedleFillStyle" at 330,690 size 95x20; Text 'NeedleFillStyle'
   Clock "NumberStyle" at 490,538 size 150x150
   TextField "Label_NumberStyle" at 490,690 size 86x20; Text 'NumberStyle'
   Clock "NumberStyle_2" at 650,538 size 150x150
   TextField "Label_NumberStyle_2" at 650,690 size 102x20; Text 'NumberStyle_2'
   Clock "SecondNeedleHeight" at 810,538 size 150x150
   TextField "Label_SecondNeedleHeight" at 810,690 size 136x20; Text 'SecondNeedleHeight'
   Button "Next" at 982,744 size 40x22; TextOff 'Text'
      on Click: ActivateScreen("P_Clock_2", 0)

screen "P_Clock_2" 1024x768
   Clock "SecondNeedleWidth" at 10,10 size 150x150
   TextField "Label_SecondNeedleWidth" at 10,162 size 132x20; Text 'SecondNeedleWidth'
   Clock "ShowTicks" at 170,10 size 150x150
   TextField "Label_ShowTicks" at 170,162 size 70x20; Text 'ShowTicks'
   Clock "TickDistance" at 330,10 size 150x150
   TextField "Label_TickDistance" at 330,162 size 84x20; Text 'TickDistance'
   Clock "TickStyle" at 490,10 size 150x150
   TextField "Label_TickStyle" at 490,162 size 61x20; Text 'TickStyle'
   Clock "TicksColor" at 650,10 size 150x150
   TextField "Label_TicksColor" at 650,162 size 68x20; Text 'TicksColor'
   Clock "UseDesignColorSchema" at 810,10 size 150x150
   TextField "Label_UseDesignColorSchema" at 810,162 size 153x20; Text 'UseDesignColorSchema'
   Button "Next" at 982,744 size 40x22; TextOff 'Text'
      on Click: ActivateScreen("P_Line_1", 0)

screen "P_IOField_1" 1024x768
   IOField "Default" at 10,10 size 100x30
   TextField "Label_Default" at 10,42 size 51x20; Text 'Default'
   IOField "AboveUpperLimitColor" at 120,10 size 100x30
   TextField "Label_AboveUpperLimitColor" at 120,42 size 147x20; Text 'AboveUpperLimitColor'
   IOField "BackColor" at 230,10 size 100x30
   TextField "Label_BackColor" at 230,42 size 67x20; Text 'BackColor'
   IOField "BackFillStyle" at 340,10 size 100x30
   TextField "Label_BackFillStyle" at 340,42 size 82x20; Text 'BackFillStyle'
   IOField "BelowLowerLimitColor" at 450,10 size 100x30
   TextField "Label_BelowLowerLimitColor" at 450,42 size 145x20; Text 'BelowLowerLimitColor'
   IOField "BorderBackColor" at 560,10 size 100x30
   TextField "Label_BorderBackColor" at 560,42 size 111x20; Text 'BorderBackColor'
   IOField "BorderColor" at 670,10 size 100x30
   TextField "Label_BorderColor" at 670,42 size 81x20; Text 'BorderColor'
   IOField "BorderWidth" at 780,10 size 100x30
   TextField "Label_BorderWidth" at 780,42 size 86x20; Text 'BorderWidth'
   IOField "BottomMargin" at 890,10 size 100x30
   TextField "Label_BottomMargin" at 890,42 size 95x20; Text 'BottomMargin'
   IOField "CornerRadius" at 10,66 size 100x30
   TextField "Label_CornerRadius" at 10,98 size 91x20; Text 'CornerRadius'
   IOField "DataFormat_3" at 120,66 size 100x30
   TextField "Label_DataFormat_3" at 120,98 size 96x20; Text 'DataFormat_3'
   IOField "EdgeStyle" at 230,66 size 100x30
   TextField "Label_EdgeStyle" at 230,98 size 68x20; Text 'EdgeStyle'
   IOField "EdgeStyle_2" at 340,66 size 100x30
   TextField "Label_EdgeStyle_2" at 340,98 size 84x20; Text 'EdgeStyle_2'
   IOField "EdgeStyle_3" at 450,66 size 100x30
   TextField "Label_EdgeStyle_3" at 450,98 size 84x20; Text 'EdgeStyle_3'
   IOField "EdgeStyle_4" at 560,66 size 100x30
   TextField "Label_EdgeStyle_4" at 560,98 size 84x20; Text 'EdgeStyle_4'
   IOField "FieldLength" at 670,66 size 100x30
   TextField "Label_FieldLength" at 670,98 size 77x20; Text 'FieldLength'
   IOField "FitToLargest" at 780,66 size 75x30
   TextField "Label_FitToLargest" at 780,98 size 84x20; Text 'FitToLargest'
   IOField "Flashing" at 890,66 size 100x30
   TextField "Label_Flashing" at 890,98 size 55x20; Text 'Flashing'
   IOField "ForeColor" at 10,122 size 100x30
   TextField "Label_ForeColor" at 10,154 size 65x20; Text 'ForeColor'
   IOField "FormatPattern" at 120,122 size 100x30; FormatPattern 99.9
   TextField "Label_FormatPattern" at 120,154 size 99x20; Text 'FormatPattern'
   IOField "HorizontalAlignment" at 230,122 size 100x30
   TextField "Label_HorizontalAlignment" at 230,154 size 135x20; Text 'HorizontalAlignment'
   IOField "HorizontalAlignment_2" at 340,122 size 100x30
   TextField "Label_HorizontalAlignment_2" at 340,154 size 151x20; Text 'HorizontalAlignment_2'
   IOField "LeftMargin" at 450,122 size 100x30
   TextField "Label_LeftMargin" at 450,154 size 74x20; Text 'LeftMargin'
   IOField "Mode" at 560,122 size 100x30
   TextField "Label_Mode" at 560,154 size 39x20; Text 'Mode'
   IOField "Mode_2" at 670,122 size 100x30
   TextField "Label_Mode_2" at 670,154 size 55x20; Text 'Mode_2'
   IOField "RightMargin" at 780,122 size 100x30
   TextField "Label_RightMargin" at 780,154 size 82x20; Text 'RightMargin'
   IOField "ShiftDecimalPoint" at 890,122 size 100x30
   TextField "Label_ShiftDecimalPoint" at 890,154 size 116x20; Text 'ShiftDecimalPoint'
   IOField "ShowLeadingZeros" at 10,178 size 100x30
   TextField "Label_ShowLeadingZeros" at 10,210 size 125x20; Text 'ShowLeadingZeros'
   IOField "TopMargin" at 120,178 size 100x30
   TextField "Label_TopMargin" at 120,210 size 71x20; Text 'TopMargin'
   IOField "Unit" at 230,178 size 100x30; Unit mm
   TextField "Label_Unit" at 230,210 size 29x20; Text 'Unit'
   IOField "UseDesignColorSchema" at 340,178 size 100x30
   TextField "Label_UseDesignColorSchema" at 340,210 size 153x20; Text 'UseDesignColorSchema'
   IOField "VerticalAlignment" at 450,178 size 100x30
   TextField "Label_VerticalAlignment" at 450,210 size 119x20; Text 'VerticalAlignment'
   IOField "VerticalAlignment_2" at 560,178 size 100x30
   TextField "Label_VerticalAlignment_2" at 560,210 size 135x20; Text 'VerticalAlignment_2'
   Button "Next" at 982,744 size 40x22; TextOff 'Text'
      on Click: ActivateScreen("P_Button_1", 0)

screen "D_Bar_1" 1024x768
   Bar "Static" at 6,4 size 40x120
   TextField "Label_Static" at 6,156 size 42x20; Text 'Static'
   Bar "A_Range" at 98,4 size 40x120
      Appearance <- "D_Range"
   TextField "Label_A_Range" at 98,156 size 63x20; Text 'A_Range'
   Bar "A_Flash" at 190,4 size 40x120
      Appearance <- "D_Range"
   TextField "Label_A_Flash" at 190,156 size 54x20; Text 'A_Flash'
   Bar "A_Bit" at 282,4 size 40x120
      Appearance <- "D_Bool"
   TextField "Label_A_Bit" at 282,156 size 39x20; Text 'A_Bit'
   Bar "A_Bits" at 374,4 size 40x120
      Appearance <- "D_Bits"
   TextField "Label_A_Bits" at 374,156 size 46x20; Text 'A_Bits'
   Bar "V_Range" at 466,4 size 40x120
      Visibility <- "D_Range"
   TextField "Label_V_Range" at 466,156 size 62x20; Text 'V_Range'
   Bar "V_Bit" at 558,4 size 40x120
      Visibility <- "D_Vis"
   TextField "Label_V_Bit" at 558,156 size 38x20; Text 'V_Bit'
   Bar "M_H" at 650,4 size 40x120
      HorizontalMovement <- "D_Pct"
   TextField "Label_M_H" at 650,156 size 32x20; Text 'M_H'
   Bar "M_V" at 742,4 size 40x120
      VerticalMovement <- "D_Pct"
   TextField "Label_M_V" at 742,156 size 32x20; Text 'M_V'
   Bar "M_D" at 834,4 size 40x120
      DiagonalMovement <- "D_Pct"
   TextField "Label_M_D" at 834,156 size 32x20; Text 'M_D'
   Bar "M_Direct" at 926,4 size 40x120
      DirectMovement <- "D_X"
      DirectMovement <- "D_Y"
   TextField "Label_M_Direct" at 926,156 size 62x20; Text 'M_Direct'
   Bar "E_Range" at 6,176 size 40x120
      ObjectEnable <- "D_Range"
   TextField "Label_E_Range" at 6,328 size 60x20; Text 'E_Range'
   Bar "E_Bit" at 98,176 size 40x120
      ObjectEnable <- "D_En"
   TextField "Label_E_Bit" at 98,328 size 36x20; Text 'E_Bit'
   Bar "PV_Pct" at 190,176 size 40x120
      ProcessValue <- "D_Pct"
   TextField "Label_PV_Pct" at 190,328 size 50x20; Text 'PV_Pct'
   Bar "PV_Real" at 282,176 size 40x120
      ProcessValue <- "D_Real"
   TextField "Label_PV_Real" at 282,328 size 57x20; Text 'PV_Real'
   Bar "PV_BarR" at 374,176 size 40x120
      ProcessValue <- "D_BarR"
   TextField "Label_PV_BarR" at 374,328 size 60x20; Text 'PV_BarR'
   Bar "PV_Pct_0_100" at 466,176 size 40x120; MinimumValue 0; MaximumValue 100
      ProcessValue <- "D_Pct"
   TextField "Label_PV_Pct_0_100" at 466,328 size 98x20; Text 'PV_Pct_0_100'
   Bar "PV_Pct_MaxMin" at 558,176 size 40x120
      ProcessValue <- "D_Pct"
      MaximumValue <- "D_Max"
      MinimumValue <- "D_Min"
   TextField "Label_PV_Pct_MaxMin" at 558,328 size 106x20; Text 'PV_Pct_MaxMin'
   IOField "State" at 4,742 size 60x22; FormatPattern 9
      ProcessValue <- "D_State"
   Button "S1" at 70,742 size 40x22; TextOff 'S1'
      on Click: "SetS1"()
   Button "S2" at 114,742 size 40x22; TextOff 'S2'
      on Click: "SetS2"()
   Button "S3" at 158,742 size 40x22; TextOff 'S3'
      on Click: "SetS3"()
   Button "S4" at 202,742 size 40x22; TextOff 'S4'
      on Click: "SetS4"()
   Button "Next" at 980,742 size 40x22; TextOff 'Next'
      on Click: ActivateScreen("D_Switch_1", 0)

screen "D_Button_1" 1024x768
   Button "Static" at 6,4 size 100x40; TextOff 'Text'
   TextField "Label_Static" at 6,76 size 42x20; Text 'Static'
   Button "A_Range" at 158,4 size 100x40; TextOff 'Text'
      Appearance <- "D_Range"
   TextField "Label_A_Range" at 158,76 size 63x20; Text 'A_Range'
   Button "A_Flash" at 310,4 size 100x40; TextOff 'Text'
      Appearance <- "D_Range"
   TextField "Label_A_Flash" at 310,76 size 54x20; Text 'A_Flash'
   Button "A_Bit" at 462,4 size 100x40; TextOff 'Text'
      Appearance <- "D_Bool"
   TextField "Label_A_Bit" at 462,76 size 39x20; Text 'A_Bit'
   Button "A_Bits" at 614,4 size 100x40; TextOff 'Text'
      Appearance <- "D_Bits"
   TextField "Label_A_Bits" at 614,76 size 46x20; Text 'A_Bits'
   Button "V_Range" at 766,4 size 100x40; TextOff 'Text'
      Visibility <- "D_Range"
   TextField "Label_V_Range" at 766,76 size 62x20; Text 'V_Range'
   Button "V_Bit" at 6,96 size 100x40; TextOff 'Text'
      Visibility <- "D_Vis"
   TextField "Label_V_Bit" at 6,168 size 38x20; Text 'V_Bit'
   Button "M_H" at 158,96 size 100x40; TextOff 'Text'
      HorizontalMovement <- "D_Pct"
   TextField "Label_M_H" at 158,168 size 32x20; Text 'M_H'
   Button "M_V" at 310,96 size 100x40; TextOff 'Text'
      VerticalMovement <- "D_Pct"
   TextField "Label_M_V" at 310,168 size 32x20; Text 'M_V'
   Button "M_D" at 462,96 size 100x40; TextOff 'Text'
      DiagonalMovement <- "D_Pct"
   TextField "Label_M_D" at 462,168 size 32x20; Text 'M_D'
   Button "M_Direct" at 614,96 size 100x40; TextOff 'Text'
      DirectMovement <- "D_X"
      DirectMovement <- "D_Y"
   TextField "Label_M_Direct" at 614,168 size 62x20; Text 'M_Direct'
   Button "E_Range" at 766,96 size 100x40; TextOff 'Text'
      ObjectEnable <- "D_Range"
   TextField "Label_E_Range" at 766,168 size 60x20; Text 'E_Range'
   Button "E_Bit" at 6,188 size 100x40; TextOff 'Text'
      ObjectEnable <- "D_En"
   TextField "Label_E_Bit" at 6,260 size 36x20; Text 'E_Bit'
   IOField "State" at 4,742 size 60x22; FormatPattern 9
      ProcessValue <- "D_State"
   Button "S1" at 70,742 size 40x22; TextOff 'S1'
      on Click: "SetS1"()
   Button "S2" at 114,742 size 40x22; TextOff 'S2'
      on Click: "SetS2"()
   Button "S3" at 158,742 size 40x22; TextOff 'S3'
      on Click: "SetS3"()
   Button "S4" at 202,742 size 40x22; TextOff 'S4'
      on Click: "SetS4"()
   Button "Next" at 980,742 size 40x22; TextOff 'Next'
      on Click: ActivateScreen("D_SymbolicIOField_1", 0)

screen "D_Circle_1" 1024x768
   TextField "Label_Static" at 6,86 size 42x20; Text 'Static'
   Circle "A_Range" at 108,4 size 50x50
      Appearance <- "D_Range"
   TextField "Label_A_Range" at 108,86 size 63x20; Text 'A_Range'
   Circle "A_Flash" at 210,4 size 50x50
      Appearance <- "D_Range"
   TextField "Label_A_Flash" at 210,86 size 54x20; Text 'A_Flash'
   Circle "A_Bit" at 312,4 size 50x50
      Appearance <- "D_Bool"
   TextField "Label_A_Bit" at 312,86 size 39x20; Text 'A_Bit'
   Circle "A_Bits" at 414,4 size 50x50
      Appearance <- "D_Bits"
   TextField "Label_A_Bits" at 414,86 size 46x20; Text 'A_Bits'
   Circle "V_Range" at 516,4 size 50x50
      Visibility <- "D_Range"
   TextField "Label_V_Range" at 516,86 size 62x20; Text 'V_Range'
   Circle "V_Bit" at 618,4 size 50x50
      Visibility <- "D_Vis"
   TextField "Label_V_Bit" at 618,86 size 38x20; Text 'V_Bit'
   Circle "M_H" at 720,4 size 50x50
      HorizontalMovement <- "D_Pct"
   TextField "Label_M_H" at 720,86 size 32x20; Text 'M_H'
   Circle "M_V" at 822,4 size 50x50
      VerticalMovement <- "D_Pct"
   TextField "Label_M_V" at 822,86 size 32x20; Text 'M_V'
   Circle "M_D" at 6,106 size 50x50
      DiagonalMovement <- "D_Pct"
   TextField "Label_M_D" at 6,188 size 32x20; Text 'M_D'
   Circle "M_Direct" at 108,106 size 50x50
      DirectMovement <- "D_X"
      DirectMovement <- "D_Y"
   TextField "Label_M_Direct" at 108,188 size 62x20; Text 'M_Direct'
   Circle "E_Range" at 210,106 size 50x50
      ObjectEnable <- "D_Range"
   TextField "Label_E_Range" at 210,188 size 60x20; Text 'E_Range'
   Circle "E_Bit" at 312,106 size 50x50
      ObjectEnable <- "D_En"
   TextField "Label_E_Bit" at 312,188 size 36x20; Text 'E_Bit'
   IOField "State" at 4,742 size 60x22; FormatPattern 9
      ProcessValue <- "D_State"
   Button "S1" at 70,742 size 40x22; TextOff 'S1'
      on Click: "SetS1"()
   Button "S2" at 114,742 size 40x22; TextOff 'S2'
      on Click: "SetS2"()
   Button "S3" at 158,742 size 40x22; TextOff 'S3'
      on Click: "SetS3"()
   Button "S4" at 202,742 size 40x22; TextOff 'S4'
      on Click: "SetS4"()
   Button "Next" at 980,742 size 40x22; TextOff 'Next'
      on Click: ActivateScreen("D_Rectangle_1", 0)

screen "D_Clock_1" 1024x768
   Clock "Static" at 6,4 size 150x150
   TextField "Label_Static" at 6,186 size 42x20; Text 'Static'
   Clock "A_Range" at 208,4 size 150x150
      Appearance <- "D_Range"
   TextField "Label_A_Range" at 208,186 size 63x20; Text 'A_Range'
   Clock "A_Flash" at 410,4 size 150x150
      Appearance <- "D_Range"
   TextField "Label_A_Flash" at 410,186 size 54x20; Text 'A_Flash'
   Clock "A_Bit" at 612,4 size 150x150
      Appearance <- "D_Bool"
   TextField "Label_A_Bit" at 612,186 size 39x20; Text 'A_Bit'
   Clock "A_Bits" at 814,4 size 150x150
      Appearance <- "D_Bits"
   TextField "Label_A_Bits" at 814,186 size 46x20; Text 'A_Bits'
   Clock "V_Range" at 6,206 size 150x150
      Visibility <- "D_Range"
   TextField "Label_V_Range" at 6,388 size 62x20; Text 'V_Range'
   Clock "V_Bit" at 208,206 size 150x150
      Visibility <- "D_Vis"
   TextField "Label_V_Bit" at 208,388 size 38x20; Text 'V_Bit'
   Clock "M_H" at 410,206 size 150x150
      HorizontalMovement <- "D_Pct"
   TextField "Label_M_H" at 410,388 size 32x20; Text 'M_H'
   Clock "M_V" at 612,206 size 150x150
      VerticalMovement <- "D_Pct"
   TextField "Label_M_V" at 612,388 size 32x20; Text 'M_V'
   Clock "M_D" at 814,206 size 150x150
      DiagonalMovement <- "D_Pct"
   TextField "Label_M_D" at 814,388 size 32x20; Text 'M_D'
   Clock "M_Direct" at 6,408 size 150x150
      DirectMovement <- "D_X"
      DirectMovement <- "D_Y"
   TextField "Label_M_Direct" at 6,590 size 62x20; Text 'M_Direct'
   Clock "E_Range" at 208,408 size 150x150
      ObjectEnable <- "D_Range"
   TextField "Label_E_Range" at 208,590 size 60x20; Text 'E_Range'
   Clock "E_Bit" at 410,408 size 150x150
      ObjectEnable <- "D_En"
   TextField "Label_E_Bit" at 410,590 size 36x20; Text 'E_Bit'
   IOField "State" at 4,742 size 60x22; FormatPattern 9
      ProcessValue <- "D_State"
   Button "S1" at 70,742 size 40x22; TextOff 'S1'
      on Click: "SetS1"()
   Button "S2" at 114,742 size 40x22; TextOff 'S2'
      on Click: "SetS2"()
   Button "S3" at 158,742 size 40x22; TextOff 'S3'
      on Click: "SetS3"()
   Button "S4" at 202,742 size 40x22; TextOff 'S4'
      on Click: "SetS4"()
   Button "Next" at 980,742 size 40x22; TextOff 'Next'
      on Click: ActivateScreen("D_Line_1", 0)

screen "D_DateTimeField_1" 1024x768
   DateTimeField "Static" at 6,4 size 189x26
   TextField "Label_Static" at 6,66 size 42x20; Text 'Static'
   DateTimeField "A_Range" at 218,4 size 189x26
      Appearance <- "D_Range"
   TextField "Label_A_Range" at 218,66 size 63x20; Text 'A_Range'
   DateTimeField "A_Flash" at 430,4 size 189x26
      Appearance <- "D_Range"
   TextField "Label_A_Flash" at 430,66 size 54x20; Text 'A_Flash'
   DateTimeField "A_Bit" at 642,4 size 189x26
      Appearance <- "D_Bool"
   TextField "Label_A_Bit" at 642,66 size 39x20; Text 'A_Bit'
   DateTimeField "A_Bits" at 6,86 size 189x26
      Appearance <- "D_Bits"
   TextField "Label_A_Bits" at 6,148 size 46x20; Text 'A_Bits'
   DateTimeField "V_Range" at 218,86 size 189x26
      Visibility <- "D_Range"
   TextField "Label_V_Range" at 218,148 size 62x20; Text 'V_Range'
   DateTimeField "V_Bit" at 430,86 size 189x26
      Visibility <- "D_Vis"
   TextField "Label_V_Bit" at 430,148 size 38x20; Text 'V_Bit'
   DateTimeField "M_H" at 642,86 size 189x26
      HorizontalMovement <- "D_Pct"
   TextField "Label_M_H" at 642,148 size 32x20; Text 'M_H'
   DateTimeField "M_V" at 6,168 size 189x26
      VerticalMovement <- "D_Pct"
   TextField "Label_M_V" at 6,230 size 32x20; Text 'M_V'
   DateTimeField "M_D" at 218,168 size 189x26
      DiagonalMovement <- "D_Pct"
   TextField "Label_M_D" at 218,230 size 32x20; Text 'M_D'
   DateTimeField "M_Direct" at 430,168 size 189x26
      DirectMovement <- "D_X"
      DirectMovement <- "D_Y"
   TextField "Label_M_Direct" at 430,230 size 62x20; Text 'M_Direct'
   DateTimeField "E_Range" at 642,168 size 189x26
      ObjectEnable <- "D_Range"
   TextField "Label_E_Range" at 642,230 size 60x20; Text 'E_Range'
   DateTimeField "E_Bit" at 6,250 size 189x26
      ObjectEnable <- "D_En"
   TextField "Label_E_Bit" at 6,312 size 36x20; Text 'E_Bit'
   DateTimeField "PV_DateTime" at 218,250 size 189x26
      ProcessValue <- "D_DateTime"
   TextField "Label_PV_DateTime" at 218,312 size 89x20; Text 'PV_DateTime'
   IOField "State" at 4,742 size 60x22; FormatPattern 9
      ProcessValue <- "D_State"
   Button "S1" at 70,742 size 40x22; TextOff 'S1'
      on Click: "SetS1"()
   Button "S2" at 114,742 size 40x22; TextOff 'S2'
      on Click: "SetS2"()
   Button "S3" at 158,742 size 40x22; TextOff 'S3'
      on Click: "SetS3"()
   Button "S4" at 202,742 size 40x22; TextOff 'S4'
      on Click: "SetS4"()
   Button "Next" at 980,742 size 40x22; TextOff 'Next'
      on Click: ActivateScreen("D_Bar_1", 0)

screen "D_Ellipse_1" 1024x768
   TextField "Label_Static" at 6,86 size 42x20; Text 'Static'
   Ellipse "A_Range" at 158,4 size 100x50
      Appearance <- "D_Range"
   TextField "Label_A_Range" at 158,86 size 63x20; Text 'A_Range'
   Ellipse "A_Flash" at 310,4 size 100x50
      Appearance <- "D_Range"
   TextField "Label_A_Flash" at 310,86 size 54x20; Text 'A_Flash'
   Ellipse "A_Bit" at 462,4 size 100x50
      Appearance <- "D_Bool"
   TextField "Label_A_Bit" at 462,86 size 39x20; Text 'A_Bit'
   Ellipse "A_Bits" at 614,4 size 100x50
      Appearance <- "D_Bits"
   TextField "Label_A_Bits" at 614,86 size 46x20; Text 'A_Bits'
   Ellipse "V_Range" at 766,4 size 100x50
      Visibility <- "D_Range"
   TextField "Label_V_Range" at 766,86 size 62x20; Text 'V_Range'
   Ellipse "V_Bit" at 6,106 size 100x50
      Visibility <- "D_Vis"
   TextField "Label_V_Bit" at 6,188 size 38x20; Text 'V_Bit'
   Ellipse "M_H" at 158,106 size 100x50
      HorizontalMovement <- "D_Pct"
   TextField "Label_M_H" at 158,188 size 32x20; Text 'M_H'
   Ellipse "M_V" at 310,106 size 100x50
      VerticalMovement <- "D_Pct"
   TextField "Label_M_V" at 310,188 size 32x20; Text 'M_V'
   Ellipse "M_D" at 462,106 size 100x50
      DiagonalMovement <- "D_Pct"
   TextField "Label_M_D" at 462,188 size 32x20; Text 'M_D'
   Ellipse "M_Direct" at 614,106 size 100x50
      DirectMovement <- "D_X"
      DirectMovement <- "D_Y"
   TextField "Label_M_Direct" at 614,188 size 62x20; Text 'M_Direct'
   Ellipse "E_Range" at 766,106 size 100x50
      ObjectEnable <- "D_Range"
   TextField "Label_E_Range" at 766,188 size 60x20; Text 'E_Range'
   Ellipse "E_Bit" at 6,208 size 100x50
      ObjectEnable <- "D_En"
   TextField "Label_E_Bit" at 6,290 size 36x20; Text 'E_Bit'
   IOField "State" at 4,742 size 60x22; FormatPattern 9
      ProcessValue <- "D_State"
   Button "S1" at 70,742 size 40x22; TextOff 'S1'
      on Click: "SetS1"()
   Button "S2" at 114,742 size 40x22; TextOff 'S2'
      on Click: "SetS2"()
   Button "S3" at 158,742 size 40x22; TextOff 'S3'
      on Click: "SetS3"()
   Button "S4" at 202,742 size 40x22; TextOff 'S4'
      on Click: "SetS4"()
   Button "Next" at 980,742 size 40x22; TextOff 'Next'
      on Click: ActivateScreen("D_Circle_1", 0)

screen "D_Gauge_1" 1024x768
   Gauge "Static" at 6,4 size 150x150; CaptionText 'SIMATIC'
   TextField "Label_Static" at 6,186 size 42x20; Text 'Static'
   Gauge "A_Range" at 208,4 size 150x150; CaptionText 'SIMATIC'
      Appearance <- "D_Range"
   TextField "Label_A_Range" at 208,186 size 63x20; Text 'A_Range'
   Gauge "A_Flash" at 410,4 size 150x150; CaptionText 'SIMATIC'
      Appearance <- "D_Range"
   TextField "Label_A_Flash" at 410,186 size 54x20; Text 'A_Flash'
   Gauge "A_Bit" at 612,4 size 150x150; CaptionText 'SIMATIC'
      Appearance <- "D_Bool"
   TextField "Label_A_Bit" at 612,186 size 39x20; Text 'A_Bit'
   Gauge "A_Bits" at 814,4 size 150x150; CaptionText 'SIMATIC'
      Appearance <- "D_Bits"
   TextField "Label_A_Bits" at 814,186 size 46x20; Text 'A_Bits'
   Gauge "V_Range" at 6,206 size 150x150; CaptionText 'SIMATIC'
      Visibility <- "D_Range"
   TextField "Label_V_Range" at 6,388 size 62x20; Text 'V_Range'
   Gauge "V_Bit" at 208,206 size 150x150; CaptionText 'SIMATIC'
      Visibility <- "D_Vis"
   TextField "Label_V_Bit" at 208,388 size 38x20; Text 'V_Bit'
   Gauge "M_H" at 410,206 size 150x150; CaptionText 'SIMATIC'
      HorizontalMovement <- "D_Pct"
   TextField "Label_M_H" at 410,388 size 32x20; Text 'M_H'
   Gauge "M_V" at 612,206 size 150x150; CaptionText 'SIMATIC'
      VerticalMovement <- "D_Pct"
   TextField "Label_M_V" at 612,388 size 32x20; Text 'M_V'
   Gauge "M_D" at 814,206 size 150x150; CaptionText 'SIMATIC'
      DiagonalMovement <- "D_Pct"
   TextField "Label_M_D" at 814,388 size 32x20; Text 'M_D'
   Gauge "M_Direct" at 6,408 size 150x150; CaptionText 'SIMATIC'
      DirectMovement <- "D_X"
      DirectMovement <- "D_Y"
   TextField "Label_M_Direct" at 6,590 size 62x20; Text 'M_Direct'
   Gauge "E_Range" at 208,408 size 150x150; CaptionText 'SIMATIC'
      ObjectEnable <- "D_Range"
   TextField "Label_E_Range" at 208,590 size 60x20; Text 'E_Range'
   Gauge "E_Bit" at 410,408 size 150x150; CaptionText 'SIMATIC'
      ObjectEnable <- "D_En"
   TextField "Label_E_Bit" at 410,590 size 36x20; Text 'E_Bit'
   Gauge "PV_Pct" at 612,408 size 150x150; CaptionText 'SIMATIC'
      ProcessValue <- "D_Pct"
   TextField "Label_PV_Pct" at 612,590 size 50x20; Text 'PV_Pct'
   Gauge "PV_Real" at 814,408 size 150x150; CaptionText 'SIMATIC'
      ProcessValue <- "D_Real"
   TextField "Label_PV_Real" at 814,590 size 57x20; Text 'PV_Real'
   IOField "State" at 4,742 size 60x22; FormatPattern 9
      ProcessValue <- "D_State"
   Button "S1" at 70,742 size 40x22; TextOff 'S1'
      on Click: "SetS1"()
   Button "S2" at 114,742 size 40x22; TextOff 'S2'
      on Click: "SetS2"()
   Button "S3" at 158,742 size 40x22; TextOff 'S3'
      on Click: "SetS3"()
   Button "S4" at 202,742 size 40x22; TextOff 'S4'
      on Click: "SetS4"()
   Button "Next" at 980,742 size 40x22; TextOff 'Next'
      on Click: ActivateScreen("D_Gauge_2", 0)

screen "D_Gauge_2" 1024x768
   Gauge "PV_Pct_MaxMin" at 6,4 size 150x150; CaptionText 'SIMATIC'
      ProcessValue <- "D_Pct"
      MaximumValue <- "D_Max"
      MinimumValue <- "D_Min"
   TextField "Label_PV_Pct_MaxMin" at 6,186 size 106x20; Text 'PV_Pct_MaxMin'
   IOField "State" at 4,742 size 60x22; FormatPattern 9
      ProcessValue <- "D_State"
   Button "S1" at 70,742 size 40x22; TextOff 'S1'
      on Click: "SetS1"()
   Button "S2" at 114,742 size 40x22; TextOff 'S2'
      on Click: "SetS2"()
   Button "S3" at 158,742 size 40x22; TextOff 'S3'
      on Click: "SetS3"()
   Button "S4" at 202,742 size 40x22; TextOff 'S4'
      on Click: "SetS4"()
   Button "Next" at 980,742 size 40x22; TextOff 'Next'
      on Click: ActivateScreen("D_Clock_1", 0)

screen "D_GraphicIOField_1" 1024x768
   GraphicIOField "Static" at 6,4 size 60x60
   TextField "Label_Static" at 6,96 size 42x20; Text 'Static'
   GraphicIOField "A_Range" at 118,4 size 60x60
      Appearance <- "D_Range"
   TextField "Label_A_Range" at 118,96 size 63x20; Text 'A_Range'
   GraphicIOField "A_Flash" at 230,4 size 60x60
      Appearance <- "D_Range"
   TextField "Label_A_Flash" at 230,96 size 54x20; Text 'A_Flash'
   GraphicIOField "A_Bit" at 342,4 size 60x60
      Appearance <- "D_Bool"
   TextField "Label_A_Bit" at 342,96 size 39x20; Text 'A_Bit'
   GraphicIOField "A_Bits" at 454,4 size 60x60
      Appearance <- "D_Bits"
   TextField "Label_A_Bits" at 454,96 size 46x20; Text 'A_Bits'
   GraphicIOField "V_Range" at 566,4 size 60x60
      Visibility <- "D_Range"
   TextField "Label_V_Range" at 566,96 size 62x20; Text 'V_Range'
   GraphicIOField "V_Bit" at 678,4 size 60x60
      Visibility <- "D_Vis"
   TextField "Label_V_Bit" at 678,96 size 38x20; Text 'V_Bit'
   GraphicIOField "M_H" at 790,4 size 60x60
      HorizontalMovement <- "D_Pct"
   TextField "Label_M_H" at 790,96 size 32x20; Text 'M_H'
   GraphicIOField "M_V" at 902,4 size 60x60
      VerticalMovement <- "D_Pct"
   TextField "Label_M_V" at 902,96 size 32x20; Text 'M_V'
   GraphicIOField "M_D" at 6,116 size 60x60
      DiagonalMovement <- "D_Pct"
   TextField "Label_M_D" at 6,208 size 32x20; Text 'M_D'
   GraphicIOField "M_Direct" at 118,116 size 60x60
      DirectMovement <- "D_X"
      DirectMovement <- "D_Y"
   TextField "Label_M_Direct" at 118,208 size 62x20; Text 'M_Direct'
   GraphicIOField "E_Range" at 230,116 size 60x60
      ObjectEnable <- "D_Range"
   TextField "Label_E_Range" at 230,208 size 60x20; Text 'E_Range'
   GraphicIOField "E_Bit" at 342,116 size 60x60
      ObjectEnable <- "D_En"
   TextField "Label_E_Bit" at 342,208 size 36x20; Text 'E_Bit'
   IOField "State" at 4,742 size 60x22; FormatPattern 9
      ProcessValue <- "D_State"
   Button "S1" at 70,742 size 40x22; TextOff 'S1'
      on Click: "SetS1"()
   Button "S2" at 114,742 size 40x22; TextOff 'S2'
      on Click: "SetS2"()
   Button "S3" at 158,742 size 40x22; TextOff 'S3'
      on Click: "SetS3"()
   Button "S4" at 202,742 size 40x22; TextOff 'S4'
      on Click: "SetS4"()
   Button "Next" at 980,742 size 40x22; TextOff 'Next'
      on Click: ActivateScreen("D_DateTimeField_1", 0)

screen "D_GraphicView_1" 1024x768
   GraphicView "Static" at 6,4 size 100x60
   TextField "Label_Static" at 6,96 size 42x20; Text 'Static'
   GraphicView "A_Range" at 158,4 size 100x60
      Appearance <- "D_Range"
   TextField "Label_A_Range" at 158,96 size 63x20; Text 'A_Range'
   GraphicView "A_Flash" at 310,4 size 100x60
      Appearance <- "D_Range"
   TextField "Label_A_Flash" at 310,96 size 54x20; Text 'A_Flash'
   GraphicView "A_Bit" at 462,4 size 100x60
      Appearance <- "D_Bool"
   TextField "Label_A_Bit" at 462,96 size 39x20; Text 'A_Bit'
   GraphicView "A_Bits" at 614,4 size 100x60
      Appearance <- "D_Bits"
   TextField "Label_A_Bits" at 614,96 size 46x20; Text 'A_Bits'
   GraphicView "V_Range" at 766,4 size 100x60
      Visibility <- "D_Range"
   TextField "Label_V_Range" at 766,96 size 62x20; Text 'V_Range'
   GraphicView "V_Bit" at 6,116 size 100x60
      Visibility <- "D_Vis"
   TextField "Label_V_Bit" at 6,208 size 38x20; Text 'V_Bit'
   GraphicView "M_H" at 158,116 size 100x60
      HorizontalMovement <- "D_Pct"
   TextField "Label_M_H" at 158,208 size 32x20; Text 'M_H'
   GraphicView "M_V" at 310,116 size 100x60
      VerticalMovement <- "D_Pct"
   TextField "Label_M_V" at 310,208 size 32x20; Text 'M_V'
   GraphicView "M_D" at 462,116 size 100x60
      DiagonalMovement <- "D_Pct"
   TextField "Label_M_D" at 462,208 size 32x20; Text 'M_D'
   GraphicView "M_Direct" at 614,116 size 100x60
      DirectMovement <- "D_X"
      DirectMovement <- "D_Y"
   TextField "Label_M_Direct" at 614,208 size 62x20; Text 'M_Direct'
   GraphicView "E_Range" at 766,116 size 100x60
      ObjectEnable <- "D_Range"
   TextField "Label_E_Range" at 766,208 size 60x20; Text 'E_Range'
   GraphicView "E_Bit" at 6,228 size 100x60
      ObjectEnable <- "D_En"
   TextField "Label_E_Bit" at 6,320 size 36x20; Text 'E_Bit'
   IOField "State" at 4,742 size 60x22; FormatPattern 9
      ProcessValue <- "D_State"
   Button "S1" at 70,742 size 40x22; TextOff 'S1'
      on Click: "SetS1"()
   Button "S2" at 114,742 size 40x22; TextOff 'S2'
      on Click: "SetS2"()
   Button "S3" at 158,742 size 40x22; TextOff 'S3'
      on Click: "SetS3"()
   Button "S4" at 202,742 size 40x22; TextOff 'S4'
      on Click: "SetS4"()
   Button "Next" at 980,742 size 40x22; TextOff 'Next'
      on Click: ActivateScreen("D_IOField_1", 0)

screen "D_IOField_1" 1024x768
   IOField "Static" at 6,4 size 100x30
   TextField "Label_Static" at 6,66 size 42x20; Text 'Static'
   IOField "A_Range" at 158,4 size 100x30
      Appearance <- "D_Range"
   TextField "Label_A_Range" at 158,66 size 63x20; Text 'A_Range'
   IOField "A_Flash" at 310,4 size 100x30
      Appearance <- "D_Range"
   TextField "Label_A_Flash" at 310,66 size 54x20; Text 'A_Flash'
   IOField "A_Bit" at 462,4 size 100x30
      Appearance <- "D_Bool"
   TextField "Label_A_Bit" at 462,66 size 39x20; Text 'A_Bit'
   IOField "A_Bits" at 614,4 size 100x30
      Appearance <- "D_Bits"
   TextField "Label_A_Bits" at 614,66 size 46x20; Text 'A_Bits'
   IOField "V_Range" at 766,4 size 100x30
      Visibility <- "D_Range"
   TextField "Label_V_Range" at 766,66 size 62x20; Text 'V_Range'
   IOField "V_Bit" at 6,86 size 100x30
      Visibility <- "D_Vis"
   TextField "Label_V_Bit" at 6,148 size 38x20; Text 'V_Bit'
   IOField "M_H" at 158,86 size 100x30
      HorizontalMovement <- "D_Pct"
   TextField "Label_M_H" at 158,148 size 32x20; Text 'M_H'
   IOField "M_V" at 310,86 size 100x30
      VerticalMovement <- "D_Pct"
   TextField "Label_M_V" at 310,148 size 32x20; Text 'M_V'
   IOField "M_D" at 462,86 size 100x30
      DiagonalMovement <- "D_Pct"
   TextField "Label_M_D" at 462,148 size 32x20; Text 'M_D'
   IOField "M_Direct" at 614,86 size 100x30
      DirectMovement <- "D_X"
      DirectMovement <- "D_Y"
   TextField "Label_M_Direct" at 614,148 size 62x20; Text 'M_Direct'
   IOField "E_Range" at 766,86 size 100x30
      ObjectEnable <- "D_Range"
   TextField "Label_E_Range" at 766,148 size 60x20; Text 'E_Range'
   IOField "E_Bit" at 6,168 size 100x30
      ObjectEnable <- "D_En"
   TextField "Label_E_Bit" at 6,230 size 36x20; Text 'E_Bit'
   IOField "PV_SInt" at 158,168 size 100x30; FormatPattern s999
      ProcessValue <- "D_SInt"
   TextField "Label_PV_SInt" at 158,230 size 56x20; Text 'PV_SInt'
   IOField "PV_Int" at 310,168 size 100x30; FormatPattern s99999
      ProcessValue <- "D_Int"
   TextField "Label_PV_Int" at 310,230 size 48x20; Text 'PV_Int'
   IOField "PV_DInt" at 462,168 size 100x30; FormatPattern s9999999999
      ProcessValue <- "D_DInt"
   TextField "Label_PV_DInt" at 462,230 size 57x20; Text 'PV_DInt'
   IOField "PV_USInt" at 614,168 size 100x30; FormatPattern 999
      ProcessValue <- "D_USInt"
   TextField "Label_PV_USInt" at 614,230 size 64x20; Text 'PV_USInt'
   IOField "PV_UInt" at 766,168 size 100x30; FormatPattern 99999
      ProcessValue <- "D_UInt"
   TextField "Label_PV_UInt" at 766,230 size 56x20; Text 'PV_UInt'
   IOField "PV_UDInt" at 6,250 size 100x30; FormatPattern 9999999999
      ProcessValue <- "D_UDInt"
   TextField "Label_PV_UDInt" at 6,312 size 65x20; Text 'PV_UDInt'
   IOField "PV_Real" at 158,250 size 100x30
      ProcessValue <- "D_Real"
   TextField "Label_PV_Real" at 158,312 size 57x20; Text 'PV_Real'
   IOField "PV_LReal" at 310,250 size 100x30
      ProcessValue <- "D_LReal"
   TextField "Label_PV_LReal" at 310,312 size 64x20; Text 'PV_LReal'
   IOField "PV_String" at 462,250 size 100x30
      ProcessValue <- "D_String"
   TextField "Label_PV_String" at 462,312 size 68x20; Text 'PV_String'
   IOField "PV_Int_Shift2" at 614,250 size 100x30; FormatPattern s99999
      ProcessValue <- "D_Int"
   TextField "Label_PV_Int_Shift2" at 614,312 size 94x20; Text 'PV_Int_Shift2'
   IOField "PV_Int_s999999" at 766,250 size 100x30; FormatPattern s999999
      ProcessValue <- "D_Int"
   TextField "Label_PV_Int_s999999" at 766,312 size 111x20; Text 'PV_Int_s999999'
   IOField "PV_Real_s9999_99" at 6,332 size 100x30; FormatPattern s9999.99
      ProcessValue <- "D_Real"
   TextField "Label_PV_Real_s9999_99" at 6,394 size 128x20; Text 'PV_Real_s9999_99'
   IOField "PV_Int_Output" at 158,332 size 100x30; FormatPattern s99999
      ProcessValue <- "D_Int"
   TextField "Label_PV_Int_Output" at 158,394 size 101x20; Text 'PV_Int_Output'
   IOField "PV_Int_s99" at 310,332 size 100x30; FormatPattern s99
      ProcessValue <- "D_Int"
   TextField "Label_PV_Int_s99" at 310,394 size 79x20; Text 'PV_Int_s99'
   IOField "State" at 4,742 size 60x22; FormatPattern 9
      ProcessValue <- "D_State"
   Button "S1" at 70,742 size 40x22; TextOff 'S1'
      on Click: "SetS1"()
   Button "S2" at 114,742 size 40x22; TextOff 'S2'
      on Click: "SetS2"()
   Button "S3" at 158,742 size 40x22; TextOff 'S3'
      on Click: "SetS3"()
   Button "S4" at 202,742 size 40x22; TextOff 'S4'
      on Click: "SetS4"()
   Button "Next" at 980,742 size 40x22; TextOff 'Next'
      on Click: ActivateScreen("D_Button_1", 0)

screen "D_Line_1" 1024x768
   TextField "Label_Static" at 6,86 size 42x20; Text 'Static'
   Line "A_Range" at 158,4 size 100x50
      Appearance <- "D_Range"
   TextField "Label_A_Range" at 158,86 size 63x20; Text 'A_Range'
   Line "A_Flash" at 310,4 size 100x50
      Appearance <- "D_Range"
   TextField "Label_A_Flash" at 310,86 size 54x20; Text 'A_Flash'
   Line "A_Bit" at 462,4 size 100x50
      Appearance <- "D_Bool"
   TextField "Label_A_Bit" at 462,86 size 39x20; Text 'A_Bit'
   Line "A_Bits" at 614,4 size 100x50
      Appearance <- "D_Bits"
   TextField "Label_A_Bits" at 614,86 size 46x20; Text 'A_Bits'
   Line "V_Range" at 766,4 size 100x50
      Visibility <- "D_Range"
   TextField "Label_V_Range" at 766,86 size 62x20; Text 'V_Range'
   Line "V_Bit" at 6,106 size 100x50
      Visibility <- "D_Vis"
   TextField "Label_V_Bit" at 6,188 size 38x20; Text 'V_Bit'
   Line "M_H" at 158,106 size 100x50
      HorizontalMovement <- "D_Pct"
   TextField "Label_M_H" at 158,188 size 32x20; Text 'M_H'
   Line "M_V" at 310,106 size 100x50
      VerticalMovement <- "D_Pct"
   TextField "Label_M_V" at 310,188 size 32x20; Text 'M_V'
   Line "M_D" at 462,106 size 100x50
      DiagonalMovement <- "D_Pct"
   TextField "Label_M_D" at 462,188 size 32x20; Text 'M_D'
   Line "M_Direct" at 614,106 size 100x50
      DirectMovement <- "D_X"
      DirectMovement <- "D_Y"
   TextField "Label_M_Direct" at 614,188 size 62x20; Text 'M_Direct'
   Line "E_Range" at 766,106 size 100x50
      ObjectEnable <- "D_Range"
   TextField "Label_E_Range" at 766,188 size 60x20; Text 'E_Range'
   Line "E_Bit" at 6,208 size 100x50
      ObjectEnable <- "D_En"
   TextField "Label_E_Bit" at 6,290 size 36x20; Text 'E_Bit'
   IOField "State" at 4,742 size 60x22; FormatPattern 9
      ProcessValue <- "D_State"
   Button "S1" at 70,742 size 40x22; TextOff 'S1'
      on Click: "SetS1"()
   Button "S2" at 114,742 size 40x22; TextOff 'S2'
      on Click: "SetS2"()
   Button "S3" at 158,742 size 40x22; TextOff 'S3'
      on Click: "SetS3"()
   Button "S4" at 202,742 size 40x22; TextOff 'S4'
      on Click: "SetS4"()
   Button "Next" at 980,742 size 40x22; TextOff 'Next'
      on Click: ActivateScreen("D_Polyline_1", 0)

screen "D_Polygon_1" 1024x768
   TextField "Label_Static" at 6,86 size 42x20; Text 'Static'
   Polygon "A_Range" at 158,4 size 100x50
      Appearance <- "D_Range"
   TextField "Label_A_Range" at 158,86 size 63x20; Text 'A_Range'
   Polygon "A_Flash" at 310,4 size 100x50
      Appearance <- "D_Range"
   TextField "Label_A_Flash" at 310,86 size 54x20; Text 'A_Flash'
   Polygon "A_Bit" at 462,4 size 100x50
      Appearance <- "D_Bool"
   TextField "Label_A_Bit" at 462,86 size 39x20; Text 'A_Bit'
   Polygon "A_Bits" at 614,4 size 100x50
      Appearance <- "D_Bits"
   TextField "Label_A_Bits" at 614,86 size 46x20; Text 'A_Bits'
   Polygon "V_Range" at 766,4 size 100x50
      Visibility <- "D_Range"
   TextField "Label_V_Range" at 766,86 size 62x20; Text 'V_Range'
   Polygon "V_Bit" at 6,106 size 100x50
      Visibility <- "D_Vis"
   TextField "Label_V_Bit" at 6,188 size 38x20; Text 'V_Bit'
   Polygon "M_H" at 158,106 size 100x50
      HorizontalMovement <- "D_Pct"
   TextField "Label_M_H" at 158,188 size 32x20; Text 'M_H'
   Polygon "M_V" at 310,106 size 100x50
      VerticalMovement <- "D_Pct"
   TextField "Label_M_V" at 310,188 size 32x20; Text 'M_V'
   Polygon "M_D" at 462,106 size 100x50
      DiagonalMovement <- "D_Pct"
   TextField "Label_M_D" at 462,188 size 32x20; Text 'M_D'
   Polygon "M_Direct" at 614,106 size 100x50
      DirectMovement <- "D_X"
      DirectMovement <- "D_Y"
   TextField "Label_M_Direct" at 614,188 size 62x20; Text 'M_Direct'
   Polygon "E_Range" at 766,106 size 100x50
      ObjectEnable <- "D_Range"
   TextField "Label_E_Range" at 766,188 size 60x20; Text 'E_Range'
   Polygon "E_Bit" at 6,208 size 100x50
      ObjectEnable <- "D_En"
   TextField "Label_E_Bit" at 6,290 size 36x20; Text 'E_Bit'
   IOField "State" at 4,742 size 60x22; FormatPattern 9
      ProcessValue <- "D_State"
   Button "S1" at 70,742 size 40x22; TextOff 'S1'
      on Click: "SetS1"()
   Button "S2" at 114,742 size 40x22; TextOff 'S2'
      on Click: "SetS2"()
   Button "S3" at 158,742 size 40x22; TextOff 'S3'
      on Click: "SetS3"()
   Button "S4" at 202,742 size 40x22; TextOff 'S4'
      on Click: "SetS4"()
   Button "Next" at 980,742 size 40x22; TextOff 'Next'
      on Click: ActivateScreen("D_Ellipse_1", 0)

screen "D_Polyline_1" 1024x768
   TextField "Label_Static" at 6,86 size 42x20; Text 'Static'
   Polyline "A_Range" at 158,4 size 100x50
      Appearance <- "D_Range"
   TextField "Label_A_Range" at 158,86 size 63x20; Text 'A_Range'
   Polyline "A_Flash" at 310,4 size 100x50
      Appearance <- "D_Range"
   TextField "Label_A_Flash" at 310,86 size 54x20; Text 'A_Flash'
   Polyline "A_Bit" at 462,4 size 100x50
      Appearance <- "D_Bool"
   TextField "Label_A_Bit" at 462,86 size 39x20; Text 'A_Bit'
   Polyline "A_Bits" at 614,4 size 100x50
      Appearance <- "D_Bits"
   TextField "Label_A_Bits" at 614,86 size 46x20; Text 'A_Bits'
   Polyline "V_Range" at 766,4 size 100x50
      Visibility <- "D_Range"
   TextField "Label_V_Range" at 766,86 size 62x20; Text 'V_Range'
   Polyline "V_Bit" at 6,106 size 100x50
      Visibility <- "D_Vis"
   TextField "Label_V_Bit" at 6,188 size 38x20; Text 'V_Bit'
   Polyline "M_H" at 158,106 size 100x50
      HorizontalMovement <- "D_Pct"
   TextField "Label_M_H" at 158,188 size 32x20; Text 'M_H'
   Polyline "M_V" at 310,106 size 100x50
      VerticalMovement <- "D_Pct"
   TextField "Label_M_V" at 310,188 size 32x20; Text 'M_V'
   Polyline "M_D" at 462,106 size 100x50
      DiagonalMovement <- "D_Pct"
   TextField "Label_M_D" at 462,188 size 32x20; Text 'M_D'
   Polyline "M_Direct" at 614,106 size 100x50
      DirectMovement <- "D_X"
      DirectMovement <- "D_Y"
   TextField "Label_M_Direct" at 614,188 size 62x20; Text 'M_Direct'
   Polyline "E_Range" at 766,106 size 100x50
      ObjectEnable <- "D_Range"
   TextField "Label_E_Range" at 766,188 size 60x20; Text 'E_Range'
   Polyline "E_Bit" at 6,208 size 100x50
      ObjectEnable <- "D_En"
   TextField "Label_E_Bit" at 6,290 size 36x20; Text 'E_Bit'
   IOField "State" at 4,742 size 60x22; FormatPattern 9
      ProcessValue <- "D_State"
   Button "S1" at 70,742 size 40x22; TextOff 'S1'
      on Click: "SetS1"()
   Button "S2" at 114,742 size 40x22; TextOff 'S2'
      on Click: "SetS2"()
   Button "S3" at 158,742 size 40x22; TextOff 'S3'
      on Click: "SetS3"()
   Button "S4" at 202,742 size 40x22; TextOff 'S4'
      on Click: "SetS4"()
   Button "Next" at 980,742 size 40x22; TextOff 'Next'
      on Click: ActivateScreen("D_Polygon_1", 0)

screen "D_Rectangle_1" 1024x768
   TextField "Label_Static" at 6,86 size 42x20; Text 'Static'
   Rectangle "A_Range" at 158,4 size 100x50
      Appearance <- "D_Range"
   TextField "Label_A_Range" at 158,86 size 63x20; Text 'A_Range'
   Rectangle "A_Flash" at 310,4 size 100x50
      Appearance <- "D_Range"
   TextField "Label_A_Flash" at 310,86 size 54x20; Text 'A_Flash'
   Rectangle "A_Bit" at 462,4 size 100x50
      Appearance <- "D_Bool"
   TextField "Label_A_Bit" at 462,86 size 39x20; Text 'A_Bit'
   Rectangle "A_Bits" at 614,4 size 100x50
      Appearance <- "D_Bits"
   TextField "Label_A_Bits" at 614,86 size 46x20; Text 'A_Bits'
   Rectangle "V_Range" at 766,4 size 100x50
      Visibility <- "D_Range"
   TextField "Label_V_Range" at 766,86 size 62x20; Text 'V_Range'
   Rectangle "V_Bit" at 6,106 size 100x50
      Visibility <- "D_Vis"
   TextField "Label_V_Bit" at 6,188 size 38x20; Text 'V_Bit'
   Rectangle "M_H" at 158,106 size 100x50
      HorizontalMovement <- "D_Pct"
   TextField "Label_M_H" at 158,188 size 32x20; Text 'M_H'
   Rectangle "M_V" at 310,106 size 100x50
      VerticalMovement <- "D_Pct"
   TextField "Label_M_V" at 310,188 size 32x20; Text 'M_V'
   Rectangle "M_D" at 462,106 size 100x50
      DiagonalMovement <- "D_Pct"
   TextField "Label_M_D" at 462,188 size 32x20; Text 'M_D'
   Rectangle "M_Direct" at 614,106 size 100x50
      DirectMovement <- "D_X"
      DirectMovement <- "D_Y"
   TextField "Label_M_Direct" at 614,188 size 62x20; Text 'M_Direct'
   Rectangle "E_Range" at 766,106 size 100x50
      ObjectEnable <- "D_Range"
   TextField "Label_E_Range" at 766,188 size 60x20; Text 'E_Range'
   Rectangle "E_Bit" at 6,208 size 100x50
      ObjectEnable <- "D_En"
   TextField "Label_E_Bit" at 6,290 size 36x20; Text 'E_Bit'
   IOField "State" at 4,742 size 60x22; FormatPattern 9
      ProcessValue <- "D_State"
   Button "S1" at 70,742 size 40x22; TextOff 'S1'
      on Click: "SetS1"()
   Button "S2" at 114,742 size 40x22; TextOff 'S2'
      on Click: "SetS2"()
   Button "S3" at 158,742 size 40x22; TextOff 'S3'
      on Click: "SetS3"()
   Button "S4" at 202,742 size 40x22; TextOff 'S4'
      on Click: "SetS4"()
   Button "Next" at 980,742 size 40x22; TextOff 'Next'
      on Click: ActivateScreen("D_TextField_1", 0)

screen "D_Slider_1" 1024x768
   Slider "Static" at 6,4 size 60x160; Caption 'SIMATIC'
   TextField "Label_Static" at 6,196 size 42x20; Text 'Static'
   Slider "A_Range" at 118,4 size 60x160; Caption 'SIMATIC'
      Appearance <- "D_Range"
   TextField "Label_A_Range" at 118,196 size 63x20; Text 'A_Range'
   Slider "A_Flash" at 230,4 size 60x160; Caption 'SIMATIC'
      Appearance <- "D_Range"
   TextField "Label_A_Flash" at 230,196 size 54x20; Text 'A_Flash'
   Slider "A_Bit" at 342,4 size 60x160; Caption 'SIMATIC'
      Appearance <- "D_Bool"
   TextField "Label_A_Bit" at 342,196 size 39x20; Text 'A_Bit'
   Slider "A_Bits" at 454,4 size 60x160; Caption 'SIMATIC'
      Appearance <- "D_Bits"
   TextField "Label_A_Bits" at 454,196 size 46x20; Text 'A_Bits'
   Slider "V_Range" at 566,4 size 60x160; Caption 'SIMATIC'
      Visibility <- "D_Range"
   TextField "Label_V_Range" at 566,196 size 62x20; Text 'V_Range'
   Slider "V_Bit" at 678,4 size 60x160; Caption 'SIMATIC'
      Visibility <- "D_Vis"
   TextField "Label_V_Bit" at 678,196 size 38x20; Text 'V_Bit'
   Slider "M_H" at 790,4 size 60x160; Caption 'SIMATIC'
      HorizontalMovement <- "D_Pct"
   TextField "Label_M_H" at 790,196 size 32x20; Text 'M_H'
   Slider "M_V" at 902,4 size 60x160; Caption 'SIMATIC'
      VerticalMovement <- "D_Pct"
   TextField "Label_M_V" at 902,196 size 32x20; Text 'M_V'
   Slider "M_D" at 6,216 size 60x160; Caption 'SIMATIC'
      DiagonalMovement <- "D_Pct"
   TextField "Label_M_D" at 6,408 size 32x20; Text 'M_D'
   Slider "M_Direct" at 118,216 size 60x160; Caption 'SIMATIC'
      DirectMovement <- "D_X"
      DirectMovement <- "D_Y"
   TextField "Label_M_Direct" at 118,408 size 62x20; Text 'M_Direct'
   Slider "E_Range" at 230,216 size 60x160; Caption 'SIMATIC'
      ObjectEnable <- "D_Range"
   TextField "Label_E_Range" at 230,408 size 60x20; Text 'E_Range'
   Slider "E_Bit" at 342,216 size 60x160; Caption 'SIMATIC'
      ObjectEnable <- "D_En"
   TextField "Label_E_Bit" at 342,408 size 36x20; Text 'E_Bit'
   Slider "PV_Pct" at 454,216 size 60x160; Caption 'SIMATIC'
      ProcessValue <- "D_Pct"
   TextField "Label_PV_Pct" at 454,408 size 50x20; Text 'PV_Pct'
   Slider "PV_Int" at 566,216 size 60x160; Caption 'SIMATIC'
      ProcessValue <- "D_Int"
   TextField "Label_PV_Int" at 566,408 size 48x20; Text 'PV_Int'
   Slider "PV_Pct_0_200" at 678,216 size 60x160; Caption 'SIMATIC'
      ProcessValue <- "D_Pct"
   TextField "Label_PV_Pct_0_200" at 678,408 size 98x20; Text 'PV_Pct_0_200'
   IOField "State" at 4,742 size 60x22; FormatPattern 9
      ProcessValue <- "D_State"
   Button "S1" at 70,742 size 40x22; TextOff 'S1'
      on Click: "SetS1"()
   Button "S2" at 114,742 size 40x22; TextOff 'S2'
      on Click: "SetS2"()
   Button "S3" at 158,742 size 40x22; TextOff 'S3'
      on Click: "SetS3"()
   Button "S4" at 202,742 size 40x22; TextOff 'S4'
      on Click: "SetS4"()
   Button "Next" at 980,742 size 40x22; TextOff 'Next'
      on Click: ActivateScreen("D_Gauge_1", 0)

screen "D_Switch_1" 1024x768
   Switch "Static" at 6,4 size 120x40; CaptionText 'Switch'; TextOff '0'; TextOn '1'
   TextField "Label_Static" at 6,76 size 42x20; Text 'Static'
   Switch "A_Range" at 178,4 size 120x40; CaptionText 'Switch'; TextOff '0'; TextOn '1'
      Appearance <- "D_Range"
   TextField "Label_A_Range" at 178,76 size 63x20; Text 'A_Range'
   Switch "A_Flash" at 350,4 size 120x40; CaptionText 'Switch'; TextOff '0'; TextOn '1'
      Appearance <- "D_Range"
   TextField "Label_A_Flash" at 350,76 size 54x20; Text 'A_Flash'
   Switch "A_Bit" at 522,4 size 120x40; CaptionText 'Switch'; TextOff '0'; TextOn '1'
      Appearance <- "D_Bool"
   TextField "Label_A_Bit" at 522,76 size 39x20; Text 'A_Bit'
   Switch "A_Bits" at 694,4 size 120x40; CaptionText 'Switch'; TextOff '0'; TextOn '1'
      Appearance <- "D_Bits"
   TextField "Label_A_Bits" at 694,76 size 46x20; Text 'A_Bits'
   Switch "V_Range" at 6,96 size 120x40; CaptionText 'Switch'; TextOff '0'; TextOn '1'
      Visibility <- "D_Range"
   TextField "Label_V_Range" at 6,168 size 62x20; Text 'V_Range'
   Switch "V_Bit" at 178,96 size 120x40; CaptionText 'Switch'; TextOff '0'; TextOn '1'
      Visibility <- "D_Vis"
   TextField "Label_V_Bit" at 178,168 size 38x20; Text 'V_Bit'
   Switch "M_H" at 350,96 size 120x40; CaptionText 'Switch'; TextOff '0'; TextOn '1'
      HorizontalMovement <- "D_Pct"
   TextField "Label_M_H" at 350,168 size 32x20; Text 'M_H'
   Switch "M_V" at 522,96 size 120x40; CaptionText 'Switch'; TextOff '0'; TextOn '1'
      VerticalMovement <- "D_Pct"
   TextField "Label_M_V" at 522,168 size 32x20; Text 'M_V'
   Switch "M_D" at 694,96 size 120x40; CaptionText 'Switch'; TextOff '0'; TextOn '1'
      DiagonalMovement <- "D_Pct"
   TextField "Label_M_D" at 694,168 size 32x20; Text 'M_D'
   Switch "M_Direct" at 6,188 size 120x40; CaptionText 'Switch'; TextOff '0'; TextOn '1'
      DirectMovement <- "D_X"
      DirectMovement <- "D_Y"
   TextField "Label_M_Direct" at 6,260 size 62x20; Text 'M_Direct'
   Switch "E_Range" at 178,188 size 120x40; CaptionText 'Switch'; TextOff '0'; TextOn '1'
      ObjectEnable <- "D_Range"
   TextField "Label_E_Range" at 178,260 size 60x20; Text 'E_Range'
   Switch "E_Bit" at 350,188 size 120x40; CaptionText 'Switch'; TextOff '0'; TextOn '1'
      ObjectEnable <- "D_En"
   TextField "Label_E_Bit" at 350,260 size 36x20; Text 'E_Bit'
   Switch "PV_Bool" at 522,188 size 120x40; CaptionText 'Switch'; TextOff '0'; TextOn '1'
      ProcessValue <- "D_Bool"
   TextField "Label_PV_Bool" at 522,260 size 56x20; Text 'PV_Bool'
   IOField "State" at 4,742 size 60x22; FormatPattern 9
      ProcessValue <- "D_State"
   Button "S1" at 70,742 size 40x22; TextOff 'S1'
      on Click: "SetS1"()
   Button "S2" at 114,742 size 40x22; TextOff 'S2'
      on Click: "SetS2"()
   Button "S3" at 158,742 size 40x22; TextOff 'S3'
      on Click: "SetS3"()
   Button "S4" at 202,742 size 40x22; TextOff 'S4'
      on Click: "SetS4"()
   Button "Next" at 980,742 size 40x22; TextOff 'Next'
      on Click: ActivateScreen("D_SymbolLibrary_1", 0)

screen "D_SymbolicIOField_1" 1024x768
   SymbolicIOField "Static" at 6,4 size 120x30; TextOff '0'; TextOn '1'
   TextField "Label_Static" at 6,66 size 42x20; Text 'Static'
   SymbolicIOField "A_Range" at 178,4 size 120x30; TextOff '0'; TextOn '1'
      Appearance <- "D_Range"
   TextField "Label_A_Range" at 178,66 size 63x20; Text 'A_Range'
   SymbolicIOField "A_Flash" at 350,4 size 120x30; TextOff '0'; TextOn '1'
      Appearance <- "D_Range"
   TextField "Label_A_Flash" at 350,66 size 54x20; Text 'A_Flash'
   SymbolicIOField "A_Bit" at 522,4 size 120x30; TextOff '0'; TextOn '1'
      Appearance <- "D_Bool"
   TextField "Label_A_Bit" at 522,66 size 39x20; Text 'A_Bit'
   SymbolicIOField "A_Bits" at 694,4 size 120x30; TextOff '0'; TextOn '1'
      Appearance <- "D_Bits"
   TextField "Label_A_Bits" at 694,66 size 46x20; Text 'A_Bits'
   SymbolicIOField "V_Range" at 6,86 size 120x30; TextOff '0'; TextOn '1'
      Visibility <- "D_Range"
   TextField "Label_V_Range" at 6,148 size 62x20; Text 'V_Range'
   SymbolicIOField "V_Bit" at 178,86 size 120x30; TextOff '0'; TextOn '1'
      Visibility <- "D_Vis"
   TextField "Label_V_Bit" at 178,148 size 38x20; Text 'V_Bit'
   SymbolicIOField "M_H" at 350,86 size 120x30; TextOff '0'; TextOn '1'
      HorizontalMovement <- "D_Pct"
   TextField "Label_M_H" at 350,148 size 32x20; Text 'M_H'
   SymbolicIOField "M_V" at 522,86 size 120x30; TextOff '0'; TextOn '1'
      VerticalMovement <- "D_Pct"
   TextField "Label_M_V" at 522,148 size 32x20; Text 'M_V'
   SymbolicIOField "M_D" at 694,86 size 120x30; TextOff '0'; TextOn '1'
      DiagonalMovement <- "D_Pct"
   TextField "Label_M_D" at 694,148 size 32x20; Text 'M_D'
   SymbolicIOField "M_Direct" at 6,168 size 120x30; TextOff '0'; TextOn '1'
      DirectMovement <- "D_X"
      DirectMovement <- "D_Y"
   TextField "Label_M_Direct" at 6,230 size 62x20; Text 'M_Direct'
   SymbolicIOField "E_Range" at 178,168 size 120x30; TextOff '0'; TextOn '1'
      ObjectEnable <- "D_Range"
   TextField "Label_E_Range" at 178,230 size 60x20; Text 'E_Range'
   SymbolicIOField "E_Bit" at 350,168 size 120x30; TextOff '0'; TextOn '1'
      ObjectEnable <- "D_En"
   TextField "Label_E_Bit" at 350,230 size 36x20; Text 'E_Bit'
   SymbolicIOField "PV_TL_Value" at 522,168 size 120x30; TextOff '0'; TextOn '1'; TextList "TL_Value"
      ProcessValue <- "D_TL"
   TextField "Label_PV_TL_Value" at 522,230 size 87x20; Text 'PV_TL_Value'
   SymbolicIOField "PV_TL_Bit" at 694,168 size 120x30; TextOff '0'; TextOn '1'; TextList "TL_Bit"
      ProcessValue <- "D_Bool"
   TextField "Label_PV_TL_Bit" at 694,230 size 68x20; Text 'PV_TL_Bit'
   SymbolicIOField "PV_TL_BitNo" at 6,250 size 120x30; TextOff '0'; TextOn '1'; TextList "TL_BitNo"
      ProcessValue <- "D_Bits"
   TextField "Label_PV_TL_BitNo" at 6,312 size 84x20; Text 'PV_TL_BitNo'
   IOField "State" at 4,742 size 60x22; FormatPattern 9
      ProcessValue <- "D_State"
   Button "S1" at 70,742 size 40x22; TextOff 'S1'
      on Click: "SetS1"()
   Button "S2" at 114,742 size 40x22; TextOff 'S2'
      on Click: "SetS2"()
   Button "S3" at 158,742 size 40x22; TextOff 'S3'
      on Click: "SetS3"()
   Button "S4" at 202,742 size 40x22; TextOff 'S4'
      on Click: "SetS4"()
   Button "Next" at 980,742 size 40x22; TextOff 'Next'
      on Click: ActivateScreen("D_GraphicIOField_1", 0)

screen "D_SymbolLibrary_1" 1024x768
   SymbolLibrary "Static" at 6,4 size 60x60
   TextField "Label_Static" at 6,96 size 42x20; Text 'Static'
   SymbolLibrary "A_Range" at 118,4 size 60x60
      Appearance <- "D_Range"
   TextField "Label_A_Range" at 118,96 size 63x20; Text 'A_Range'
   SymbolLibrary "A_Flash" at 230,4 size 60x60
      Appearance <- "D_Range"
   TextField "Label_A_Flash" at 230,96 size 54x20; Text 'A_Flash'
   SymbolLibrary "A_Bit" at 342,4 size 60x60
      Appearance <- "D_Bool"
   TextField "Label_A_Bit" at 342,96 size 39x20; Text 'A_Bit'
   SymbolLibrary "A_Bits" at 454,4 size 60x60
      Appearance <- "D_Bits"
   TextField "Label_A_Bits" at 454,96 size 46x20; Text 'A_Bits'
   SymbolLibrary "V_Range" at 566,4 size 60x60
      Visibility <- "D_Range"
   TextField "Label_V_Range" at 566,96 size 62x20; Text 'V_Range'
   SymbolLibrary "V_Bit" at 678,4 size 60x60
      Visibility <- "D_Vis"
   TextField "Label_V_Bit" at 678,96 size 38x20; Text 'V_Bit'
   SymbolLibrary "M_H" at 790,4 size 60x60
      HorizontalMovement <- "D_Pct"
   TextField "Label_M_H" at 790,96 size 32x20; Text 'M_H'
   SymbolLibrary "M_V" at 902,4 size 60x60
      VerticalMovement <- "D_Pct"
   TextField "Label_M_V" at 902,96 size 32x20; Text 'M_V'
   SymbolLibrary "M_D" at 6,116 size 60x60
      DiagonalMovement <- "D_Pct"
   TextField "Label_M_D" at 6,208 size 32x20; Text 'M_D'
   SymbolLibrary "M_Direct" at 118,116 size 60x60
      DirectMovement <- "D_X"
      DirectMovement <- "D_Y"
   TextField "Label_M_Direct" at 118,208 size 62x20; Text 'M_Direct'
   SymbolLibrary "E_Range" at 230,116 size 60x60
      ObjectEnable <- "D_Range"
   TextField "Label_E_Range" at 230,208 size 60x20; Text 'E_Range'
   SymbolLibrary "E_Bit" at 342,116 size 60x60
      ObjectEnable <- "D_En"
   TextField "Label_E_Bit" at 342,208 size 36x20; Text 'E_Bit'
   SymbolLibrary "PV_Pct" at 454,116 size 60x60
      ProcessValue <- "D_Pct"
   TextField "Label_PV_Pct" at 454,208 size 50x20; Text 'PV_Pct'
   IOField "State" at 4,742 size 60x22; FormatPattern 9
      ProcessValue <- "D_State"
   Button "S1" at 70,742 size 40x22; TextOff 'S1'
      on Click: "SetS1"()
   Button "S2" at 114,742 size 40x22; TextOff 'S2'
      on Click: "SetS2"()
   Button "S3" at 158,742 size 40x22; TextOff 'S3'
      on Click: "SetS3"()
   Button "S4" at 202,742 size 40x22; TextOff 'S4'
      on Click: "SetS4"()
   Button "Next" at 980,742 size 40x22; TextOff 'Next'
      on Click: ActivateScreen("D_Slider_1", 0)

screen "D_TextField_1" 1024x768
   TextField "Static" at 6,4 size 32x20; Text 'Text'
   TextField "Label_Static" at 6,66 size 42x20; Text 'Static'
   TextField "A_Range" at 158,4 size 32x20; Text 'Text'
      Appearance <- "D_Range"
   TextField "Label_A_Range" at 158,66 size 63x20; Text 'A_Range'
   TextField "A_Flash" at 310,4 size 32x20; Text 'Text'
      Appearance <- "D_Range"
   TextField "Label_A_Flash" at 310,66 size 54x20; Text 'A_Flash'
   TextField "A_Bit" at 462,4 size 32x20; Text 'Text'
      Appearance <- "D_Bool"
   TextField "Label_A_Bit" at 462,66 size 39x20; Text 'A_Bit'
   TextField "A_Bits" at 614,4 size 32x20; Text 'Text'
      Appearance <- "D_Bits"
   TextField "Label_A_Bits" at 614,66 size 46x20; Text 'A_Bits'
   TextField "V_Range" at 766,4 size 32x20; Text 'Text'
      Visibility <- "D_Range"
   TextField "Label_V_Range" at 766,66 size 62x20; Text 'V_Range'
   TextField "V_Bit" at 6,86 size 32x20; Text 'Text'
      Visibility <- "D_Vis"
   TextField "Label_V_Bit" at 6,148 size 38x20; Text 'V_Bit'
   TextField "M_H" at 158,86 size 32x20; Text 'Text'
      HorizontalMovement <- "D_Pct"
   TextField "Label_M_H" at 158,148 size 32x20; Text 'M_H'
   TextField "M_V" at 310,86 size 32x20; Text 'Text'
      VerticalMovement <- "D_Pct"
   TextField "Label_M_V" at 310,148 size 32x20; Text 'M_V'
   TextField "M_D" at 462,86 size 32x20; Text 'Text'
      DiagonalMovement <- "D_Pct"
   TextField "Label_M_D" at 462,148 size 32x20; Text 'M_D'
   TextField "M_Direct" at 614,86 size 32x20; Text 'Text'
      DirectMovement <- "D_X"
      DirectMovement <- "D_Y"
   TextField "Label_M_Direct" at 614,148 size 62x20; Text 'M_Direct'
   TextField "E_Range" at 766,86 size 32x20; Text 'Text'
      ObjectEnable <- "D_Range"
   TextField "Label_E_Range" at 766,148 size 60x20; Text 'E_Range'
   TextField "E_Bit" at 6,168 size 32x20; Text 'Text'
      ObjectEnable <- "D_En"
   TextField "Label_E_Bit" at 6,230 size 36x20; Text 'E_Bit'
   IOField "State" at 4,742 size 60x22; FormatPattern 9
      ProcessValue <- "D_State"
   Button "S1" at 70,742 size 40x22; TextOff 'S1'
      on Click: "SetS1"()
   Button "S2" at 114,742 size 40x22; TextOff 'S2'
      on Click: "SetS2"()
   Button "S3" at 158,742 size 40x22; TextOff 'S3'
      on Click: "SetS3"()
   Button "S4" at 202,742 size 40x22; TextOff 'S4'
      on Click: "SetS4"()
   Button "Next" at 980,742 size 40x22; TextOff 'Next'
      on Click: ActivateScreen("D_GraphicView_1", 0)

screen "C5_Buttons" 1024x768, template "T_C05"
   Button "Btn_Text" at 6,40 size 120x50; TextOff 'Btn_Text off'; TextOn 'Btn_Text on'
   TextField "Label_Btn_Text" at 6,92 size 62x20; Text 'Btn_Text'
   Button "Btn_Graphic" at 182,40 size 120x90; TextOff 'Btn_Graphic off'; TextOn 'Btn_Graphic on'; PictureOff "G_PNG"; PictureOn "G_JPG"
   TextField "Label_Btn_Graphic" at 182,132 size 82x20; Text 'Btn_Graphic'
   Button "Btn_GraphicAndText" at 358,40 size 120x90; TextOff 'Btn_GraphicAndText off'; TextOn 'Btn_GraphicAndText on'; PictureOff "G_SVG"; PictureOn "G_EMF"
   TextField "Label_Btn_GraphicAndText" at 358,132 size 136x20; Text 'Btn_GraphicAndText'
   Button "Btn_TextList" at 534,40 size 160x50; TextOff 'Btn_TextList off'; TextOn 'Btn_TextList on'; TextList "TL_Value"
      ProcessValue <- "D_TL"
   TextField "Label_Btn_TextList" at 534,92 size 85x20; Text 'Btn_TextList'
   Button "Btn_GraphicList" at 710,40 size 120x90; TextOff 'Btn_GraphicList off'; TextOn 'Btn_GraphicList on'; PictureList "GL_Value"
      ProcessValue <- "D_TL"
   TextField "Label_Btn_GraphicList" at 710,132 size 105x20; Text 'Btn_GraphicList'
   Button "Btn_Invisible" at 6,152 size 120x50; TextOff 'Btn_Invisible off'; TextOn 'Btn_Invisible on'
   TextField "Label_Btn_Invisible" at 6,204 size 87x20; Text 'Btn_Invisible'
   Switch "Sw_Switch" at 182,152 size 120x40; CaptionText 'Switch'; TextOff '0'; TextOn '1'
      ProcessValue <- "D_Bool"
   TextField "Label_Sw_Switch" at 182,194 size 74x20; Text 'Sw_Switch'
   Switch "Sw_Text" at 358,152 size 120x40; CaptionText 'Switch'; TextOff 'Sw_Text off'; TextOn 'Sw_Text on'
      ProcessValue <- "D_Bool"
   TextField "Label_Sw_Text" at 358,194 size 59x20; Text 'Sw_Text'
   Switch "Sw_Graphic" at 534,152 size 120x90; CaptionText 'Switch'; TextOff '0'; TextOn '1'; PictureOff "G_BMP"; PictureOn "G_GIF"
      ProcessValue <- "D_Bool"
   TextField "Label_Sw_Graphic" at 534,244 size 79x20; Text 'Sw_Graphic'
   IOField "State" at 4,742 size 60x22; FormatPattern 9
      ProcessValue <- "D_State"
   Button "S1" at 70,742 size 40x22; TextOff 'S1'
      on Click: "SetS1"()
   Button "S2" at 114,742 size 40x22; TextOff 'S2'
      on Click: "SetS2"()
   Button "S3" at 158,742 size 40x22; TextOff 'S3'
      on Click: "SetS3"()
   Button "S4" at 202,742 size 40x22; TextOff 'S4'
      on Click: "SetS4"()
   Button "Next" at 980,742 size 40x22; TextOff 'Next'
      on Click: ActivateScreen("C5_Structure", 0)

screen "C5_GraphicView_1" 1024x768, template "T_C05"
   GraphicView "GV_PNG" at 6,40 size 120x80; Picture "G_PNG"
   TextField "Label_GV_PNG" at 6,122 size 53x20; Text 'GV_PNG'
   GraphicView "GV_JPG" at 142,40 size 120x80; Picture "G_JPG"
   TextField "Label_GV_JPG" at 142,122 size 51x20; Text 'GV_JPG'
   GraphicView "GV_BMP" at 278,40 size 120x80; Picture "G_BMP"
   TextField "Label_GV_BMP" at 278,122 size 56x20; Text 'GV_BMP'
   GraphicView "GV_GIF" at 414,40 size 120x80; Picture "G_GIF"
   TextField "Label_GV_GIF" at 414,122 size 48x20; Text 'GV_GIF'
   GraphicView "GV_TIF" at 550,40 size 120x80; Picture "G_TIF"
   TextField "Label_GV_TIF" at 550,122 size 47x20; Text 'GV_TIF'
   GraphicView "GV_EMF" at 686,40 size 120x80; Picture "G_EMF"
   TextField "Label_GV_EMF" at 686,122 size 53x20; Text 'GV_EMF'
   GraphicView "GV_WMF" at 822,40 size 120x80; Picture "G_WMF"
   TextField "Label_GV_WMF" at 822,122 size 59x20; Text 'GV_WMF'
   GraphicView "GV_SVG" at 6,142 size 120x80; Picture "G_SVG"
   TextField "Label_GV_SVG" at 6,224 size 54x20; Text 'GV_SVG'
   GraphicView "GV_TALL" at 142,142 size 120x80; Picture "G_TALL"
   TextField "Label_GV_TALL" at 142,224 size 60x20; Text 'GV_TALL'
   GraphicView "GV_WIDE" at 278,142 size 120x80; Picture "G_WIDE"
   TextField "Label_GV_WIDE" at 278,224 size 63x20; Text 'GV_WIDE'
   IOField "State" at 4,742 size 60x22; FormatPattern 9
      ProcessValue <- "D_State"
   Button "S1" at 70,742 size 40x22; TextOff 'S1'
      on Click: "SetS1"()
   Button "S2" at 114,742 size 40x22; TextOff 'S2'
      on Click: "SetS2"()
   Button "S3" at 158,742 size 40x22; TextOff 'S3'
      on Click: "SetS3"()
   Button "S4" at 202,742 size 40x22; TextOff 'S4'
      on Click: "SetS4"()
   Button "Next" at 980,742 size 40x22; TextOff 'Next'
      on Click: ActivateScreen("C5_GraphicView_2", 0)

